  movel([0.215229, -1.349679, -2.570749, -0.791960, 1.570796, 1.786025],accel_mss,speed_ms,0,blend_radius_m)
  movel([0.214975, -1.350752, -2.570030, -0.791607, 1.570796, 1.785771],accel_mss,speed_ms,0,blend_radius_m)
  movel([0.216793, -1.350982, -2.569876, -0.791531, 1.570796, 1.787589],accel_mss,speed_ms,0,blend_radius_m)
  movel([0.217496, -1.351072, -2.569815, -0.791501, 1.570796, 1.788292],accel_mss,speed_ms,0,blend_radius_m)
  movel([0.218102, -1.351157, -2.569759, -0.791474, 1.570796, 1.788899],accel_mss,speed_ms,0,blend_radius_m)
  movel([0.218626, -1.351233, -2.569708, -0.791449, 1.570796, 1.789422],accel_mss,speed_ms,0,blend_radius_m)
  movel([0.218706, -1.351253, -2.569694, -0.791442, 1.570796, 1.789502],accel_mss,speed_ms,0,blend_radius_m)
  movel([0.218724, -1.351267, -2.569684, -0.791437, 1.570796, 1.789520],accel_mss,speed_ms,0,blend_radius_m)
  movel([0.218733, -1.351290, -2.569669, -0.791430, 1.570796, 1.789529],accel_mss,speed_ms,0,blend_radius_m)
  movel([0.218734, -1.351316, -2.569652, -0.791421, 1.570796, 1.789530],accel_mss,speed_ms,0,blend_radius_m)
  movel([0.218624, -1.351824, -2.569310, -0.791255, 1.570796, 1.789420],accel_mss,speed_ms,0,blend_radius_m)
  movel([0.218549, -1.352134, -2.569101, -0.791153, 1.570796, 1.789345],accel_mss,speed_ms,0,blend_radius_m)
  movel([0.218472, -1.352445, -2.568892, -0.791052, 1.570796, 1.789269],accel_mss,speed_ms,0,blend_radius_m)
  movel([0.218266, -1.353205, -2.568380, -0.790804, 1.570796, 1.789063],accel_mss,speed_ms,0,blend_radius_m)
  movel([0.216610, -1.359807, -2.563898, -0.788684, 1.570796, 1.787406],accel_mss,speed_ms,0,blend_radius_m)
  movel([0.214499, -1.360772, -2.563238, -0.788379, 1.570796, 1.785296],accel_mss,speed_ms,0,blend_radius_m)
  movel([0.212391, -1.361738, -2.562575, -0.788076, 1.570796, 1.783188],accel_mss,speed_ms,0,blend_radius_m)
  movel([0.212109, -1.362945, -2.561746, -0.787698, 1.570796, 1.782905],accel_mss,speed_ms,0,blend_radius_m)
  movel([0.211827, -1.364150, -2.560916, -0.787322, 1.570796, 1.782623],accel_mss,speed_ms,0,blend_radius_m)
  movel([0.210167, -1.364988, -2.560338, -0.787063, 1.570796, 1.780964],accel_mss,speed_ms,0,blend_radius_m)
  movel([0.208509, -1.365829, -2.559757, -0.786803, 1.570796, 1.779305],accel_mss,speed_ms,0,blend_radius_m)
  movel([0.208371, -1.366429, -2.559341, -0.786619, 1.570796, 1.779167],accel_mss,speed_ms,0,blend_radius_m)
  movel([0.208233, -1.367028, -2.558926, -0.786435, 1.570796, 1.779029],accel_mss,speed_ms,0,blend_radius_m)
  speed_ms = 0.003
  movel([0.208233, -1.370183, -2.560451, -0.781755, 1.570796, 1.779029],accel_mss,speed_ms,0,blend_radius_m)
  speed_ms = 0.007
  movel([0.192461, -1.373239, -2.558315, -0.780834, 1.570796, 1.763257],accel_mss,speed_ms,0,blend_radius_m)
  movel([0.176700, -1.376487, -2.556031, -0.779871, 1.570796, 1.747496],accel_mss,speed_ms,0,blend_radius_m)
  movel([0.177720, -1.375452, -2.556761, -0.780176, 1.570796, 1.748516],accel_mss,speed_ms,0,blend_radius_m)
  movel([0.178177, -1.374979, -2.557093, -0.780317, 1.570796, 1.748973],accel_mss,speed_ms,0,blend_radius_m)
  movel([0.178623, -1.374493, -2.557435, -0.780461, 1.570796, 1.749419],accel_mss,speed_ms,0,blend_radius_m)
  movel([0.179054, -1.374002, -2.557780, -0.780607, 1.570796, 1.749850],accel_mss,speed_ms,0,blend_radius_m)
  movel([0.179470, -1.373501, -2.558132, -0.780756, 1.570796, 1.750267],accel_mss,speed_ms,0,blend_radius_m)
  movel([0.179870, -1.372995, -2.558487, -0.780908, 1.570796, 1.750666],accel_mss,speed_ms,0,blend_radius_m)
  movel([0.180257, -1.372480, -2.558847, -0.781062, 1.570796, 1.751054],accel_mss,speed_ms,0,blend_radius_m)
  movel([0.180628, -1.371960, -2.559211, -0.781218, 1.570796, 1.751424],accel_mss,speed_ms,0,blend_radius_m)
  movel([0.180979, -1.371442, -2.559573, -0.781374, 1.570796, 1.751775],accel_mss,speed_ms,0,blend_radius_m)
  movel([0.181310, -1.370919, -2.559938, -0.781532, 1.570796, 1.752107],accel_mss,speed_ms,0,blend_radius_m)
  movel([0.181624, -1.370393, -2.560304, -0.781691, 1.570796, 1.752420],accel_mss,speed_ms,0,blend_radius_m)
  movel([0.181922, -1.369862, -2.560675, -0.781852, 1.570796, 1.752718],accel_mss,speed_ms,0,blend_radius_m)
  movel([0.182200, -1.369330, -2.561045, -0.782014, 1.570796, 1.752996],accel_mss,speed_ms,0,blend_radius_m)
  movel([0.182457, -1.368796, -2.561416, -0.782177, 1.570796, 1.753253],accel_mss,speed_ms,0,blend_radius_m)
  movel([0.182698, -1.368260, -2.561788, -0.782341, 1.570796, 1.753494],accel_mss,speed_ms,0,blend_radius_m)
  movel([0.182918, -1.367722, -2.562161, -0.782505, 1.570796, 1.753714],accel_mss,speed_ms,0,blend_radius_m)
  movel([0.183120, -1.367184, -2.562534, -0.782671, 1.570796, 1.753916],accel_mss,speed_ms,0,blend_radius_m)
  movel([0.183301, -1.366645, -2.562907, -0.782837, 1.570796, 1.754097],accel_mss,speed_ms,0,blend_radius_m)
  movel([0.183460, -1.366110, -2.563277, -0.783002, 1.570796, 1.754256],accel_mss,speed_ms,0,blend_radius_m)
  movel([0.183600, -1.365577, -2.563645, -0.783167, 1.570796, 1.754396],accel_mss,speed_ms,0,blend_radius_m)
  movel([0.183717, -1.365048, -2.564010, -0.783331, 1.570796, 1.754514],accel_mss,speed_ms,0,blend_radius_m)
  movel([0.183813, -1.364523, -2.564372, -0.783494, 1.570796, 1.754609],accel_mss,speed_ms,0,blend_radius_m)
  movel([0.183892, -1.363989, -2.564740, -0.783660, 1.570796, 1.754688],accel_mss,speed_ms,0,blend_radius_m)
  movel([0.183948, -1.363461, -2.565103, -0.783825, 1.570796, 1.754744],accel_mss,speed_ms,0,blend_radius_m)
  movel([0.183986, -1.362939, -2.565462, -0.783988, 1.570796, 1.754782],accel_mss,speed_ms,0,blend_radius_m)
  movel([0.184002, -1.362423, -2.565816, -0.784150, 1.570796, 1.754798],accel_mss,speed_ms,0,blend_radius_m)
  movel([0.183994, -1.361916, -2.566163, -0.784310, 1.570796, 1.754790],accel_mss,speed_ms,0,blend_radius_m)
  movel([0.183968, -1.361415, -2.566506, -0.784468, 1.570796, 1.754765],accel_mss,speed_ms,0,blend_radius_m)
  movel([0.183922, -1.360922, -2.566843, -0.784623, 1.570796, 1.754718],accel_mss,speed_ms,0,blend_radius_m)
  movel([0.183841, -1.360413, -2.567192, -0.784784, 1.570796, 1.754637],accel_mss,speed_ms,0,blend_radius_m)
  movel([0.183722, -1.359924, -2.567525, -0.784939, 1.570796, 1.754519],accel_mss,speed_ms,0,blend_radius_m)
  movel([0.183540, -1.359341, -2.567923, -0.785125, 1.570796, 1.754336],accel_mss,speed_ms,0,blend_radius_m)
  movel([0.183332, -1.358771, -2.568312, -0.785307, 1.570796, 1.754129],accel_mss,speed_ms,0,blend_radius_m)
  movel([0.183103, -1.358222, -2.568685, -0.785482, 1.570796, 1.753900],accel_mss,speed_ms,0,blend_radius_m)
  movel([0.182850, -1.357690, -2.569047, -0.785652, 1.570796, 1.753646],accel_mss,speed_ms,0,blend_radius_m)
  movel([0.182624, -1.357296, -2.569314, -0.785779, 1.570796, 1.753421],accel_mss,speed_ms,0,blend_radius_m)
  movel([0.182360, -1.356931, -2.569562, -0.785896, 1.570796, 1.753156],accel_mss,speed_ms,0,blend_radius_m)
  movel([0.181837, -1.356285, -2.570000, -0.786104, 1.570796, 1.752633],accel_mss,speed_ms,0,blend_radius_m)
  movel([0.183063, -1.355949, -2.570227, -0.786213, 1.570796, 1.753859],accel_mss,speed_ms,0,blend_radius_m)
  movel([0.183512, -1.355833, -2.570306, -0.786250, 1.570796, 1.754308],accel_mss,speed_ms,0,blend_radius_m)
  movel([0.183955, -1.355730, -2.570375, -0.786283, 1.570796, 1.754752],accel_mss,speed_ms,0,blend_radius_m)
  movel([0.188162, -1.354804, -2.571002, -0.786583, 1.570796, 1.758958],accel_mss,speed_ms,0,blend_radius_m)
  movel([0.193088, -1.353747, -2.571715, -0.786927, 1.570796, 1.763885],accel_mss,speed_ms,0,blend_radius_m)
  movel([0.198699, -1.352579, -2.572501, -0.787309, 1.570796, 1.769495],accel_mss,speed_ms,0,blend_radius_m)
  movel([0.213116, -1.349701, -2.574430, -0.788258, 1.570796, 1.783912],accel_mss,speed_ms,0,blend_radius_m)
  movel([0.212938, -1.350458, -2.573924, -0.788007, 1.570796, 1.783735],accel_mss,speed_ms,0,blend_radius_m)
  movel([0.212761, -1.351214, -2.573418, -0.787758, 1.570796, 1.783557],accel_mss,speed_ms,0,blend_radius_m)
  movel([0.213243, -1.351323, -2.573344, -0.787721, 1.570796, 1.784040],accel_mss,speed_ms,0,blend_radius_m)
  movel([0.215483, -1.351799, -2.573025, -0.787565, 1.570796, 1.786280],accel_mss,speed_ms,0,blend_radius_m)
  movel([0.215229, -1.352874, -2.572303, -0.787212, 1.570796, 1.786025],accel_mss,speed_ms,0,blend_radius_m)
  movel([0.214975, -1.353945, -2.571582, -0.786863, 1.570796, 1.785771],accel_mss,speed_ms,0,blend_radius_m)
  movel([0.216793, -1.354174, -2.571427, -0.786788, 1.570796, 1.787589],accel_mss,speed_ms,0,blend_radius_m)
  movel([0.217496, -1.354264, -2.571366, -0.786759, 1.570796, 1.788292],accel_mss,speed_ms,0,blend_radius_m)
  movel([0.218102, -1.354348, -2.571309, -0.786732, 1.570796, 1.788899],accel_mss,speed_ms,0,blend_radius_m)
  movel([0.218626, -1.354424, -2.571258, -0.786707, 1.570796, 1.789422],accel_mss,speed_ms,0,blend_radius_m)
  movel([0.218706, -1.354444, -2.571245, -0.786700, 1.570796, 1.789502],accel_mss,speed_ms,0,blend_radius_m)
  movel([0.218724, -1.354458, -2.571235, -0.786696, 1.570796, 1.789520],accel_mss,speed_ms,0,blend_radius_m)
  movel([0.218733, -1.354481, -2.571220, -0.786688, 1.570796, 1.789529],accel_mss,speed_ms,0,blend_radius_m)
  movel([0.218734, -1.354507, -2.571202, -0.786680, 1.570796, 1.789530],accel_mss,speed_ms,0,blend_radius_m)
  movel([0.218624, -1.355014, -2.570860, -0.786515, 1.570796, 1.789420],accel_mss,speed_ms,0,blend_radius_m)
  movel([0.218549, -1.355323, -2.570651, -0.786415, 1.570796, 1.789345],accel_mss,speed_ms,0,blend_radius_m)
  movel([0.218472, -1.355633, -2.570441, -0.786315, 1.570796, 1.789269],accel_mss,speed_ms,0,blend_radius_m)
  movel([0.218266, -1.356391, -2.569928, -0.786070, 1.570796, 1.789063],accel_mss,speed_ms,0,blend_radius_m)
  movel([0.216610, -1.362978, -2.565435, -0.783976, 1.570796, 1.787406],accel_mss,speed_ms,0,blend_radius_m)
  movel([0.214499, -1.363941, -2.564773, -0.783675, 1.570796, 1.785296],accel_mss,speed_ms,0,blend_radius_m)
  movel([0.212391, -1.364905, -2.564109, -0.783375, 1.570796, 1.783188],accel_mss,speed_ms,0,blend_radius_m)
  movel([0.212109, -1.366109, -2.563278, -0.783002, 1.570796, 1.782905],accel_mss,speed_ms,0,blend_radius_m)
  movel([0.211827, -1.367312, -2.562446, -0.782631, 1.570796, 1.782623],accel_mss,speed_ms,0,blend_radius_m)
  movel([0.210167, -1.368148, -2.561866, -0.782375, 1.570796, 1.780964],accel_mss,speed_ms,0,blend_radius_m)
  movel([0.208509, -1.368986, -2.561284, -0.782119, 1.570796, 1.779305],accel_mss,speed_ms,0,blend_radius_m)
  movel([0.208371, -1.369585, -2.560868, -0.781937, 1.570796, 1.779167],accel_mss,speed_ms,0,blend_radius_m)
  movel([0.208233, -1.370183, -2.560451, -0.781755, 1.570796, 1.779029],accel_mss,speed_ms,0,blend_radius_m)
  speed_ms = 0.003
  movel([0.208233, -1.357697, -2.554302, -0.800390, 1.570796, 1.779029],accel_mss,speed_ms,0,blend_radius_m)
  speed_ms = 0.01
  movel([0.208233, -1.333772, -2.541623, -0.836993, 1.570796, 1.779029],accel_mss,speed_ms,0,blend_radius_m)
  movel([0.180390, -1.333590, -2.541744, -0.837055, 1.570796, 1.751186],accel_mss,speed_ms,0,blend_radius_m)
  movel([0.180390, -1.357518, -2.554425, -0.800447, 1.570796, 1.751186],accel_mss,speed_ms,0,blend_radius_m)
  speed_ms = 0.003
  movel([0.180390, -1.366850, -2.559050, -0.786489, 1.570796, 1.751186],accel_mss,speed_ms,0,blend_radius_m)
  speed_ms = 0.007
  movel([0.180139, -1.367279, -2.558752, -0.786358, 1.570796, 1.750935],accel_mss,speed_ms,0,blend_radius_m)
  movel([0.179877, -1.367706, -2.558456, -0.786227, 1.570796, 1.750673],accel_mss,speed_ms,0,blend_radius_m)
  movel([0.179604, -1.368128, -2.558163, -0.786098, 1.570796, 1.750400],accel_mss,speed_ms,0,blend_radius_m)
  movel([0.179318, -1.368547, -2.557871, -0.785971, 1.570796, 1.750115],accel_mss,speed_ms,0,blend_radius_m)
  movel([0.179021, -1.368963, -2.557582, -0.785844, 1.570796, 1.749818],accel_mss,speed_ms,0,blend_radius_m)
  movel([0.178714, -1.369376, -2.557294, -0.785719, 1.570796, 1.749510],accel_mss,speed_ms,0,blend_radius_m)
  movel([0.178399, -1.369774, -2.557017, -0.785598, 1.570796, 1.749196],accel_mss,speed_ms,0,blend_radius_m)
  movel([0.178077, -1.370168, -2.556742, -0.785479, 1.570796, 1.748873],accel_mss,speed_ms,0,blend_radius_m)
  movel([0.177744, -1.370558, -2.556470, -0.785361, 1.570796, 1.748540],accel_mss,speed_ms,0,blend_radius_m)
  movel([0.177401, -1.370941, -2.556202, -0.785246, 1.570796, 1.748197],accel_mss,speed_ms,0,blend_radius_m)
  movel([0.177050, -1.371317, -2.555939, -0.785133, 1.570796, 1.747846],accel_mss,speed_ms,0,blend_radius_m)
  movel([0.176686, -1.371687, -2.555680, -0.785022, 1.570796, 1.747483],accel_mss,speed_ms,0,blend_radius_m)
  movel([0.176338, -1.372028, -2.555441, -0.784919, 1.570796, 1.747134],accel_mss,speed_ms,0,blend_radius_m)
  movel([0.175979, -1.372363, -2.555207, -0.784819, 1.570796, 1.746776],accel_mss,speed_ms,0,blend_radius_m)
  movel([0.175611, -1.372687, -2.554979, -0.784722, 1.570796, 1.746408],accel_mss,speed_ms,0,blend_radius_m)
  movel([0.175233, -1.373005, -2.554756, -0.784627, 1.570796, 1.746029],accel_mss,speed_ms,0,blend_radius_m)
  movel([0.174850, -1.373312, -2.554541, -0.784536, 1.570796, 1.745646],accel_mss,speed_ms,0,blend_radius_m)
  movel([0.174458, -1.373609, -2.554332, -0.784447, 1.570796, 1.745254],accel_mss,speed_ms,0,blend_radius_m)
  movel([0.174093, -1.373873, -2.554147, -0.784369, 1.570796, 1.744889],accel_mss,speed_ms,0,blend_radius_m)
  movel([0.173720, -1.374131, -2.553966, -0.784293, 1.570796, 1.744516],accel_mss,speed_ms,0,blend_radius_m)
  movel([0.173344, -1.374381, -2.553790, -0.784219, 1.570796, 1.744141],accel_mss,speed_ms,0,blend_radius_m)
  movel([0.172966, -1.374620, -2.553621, -0.784148, 1.570796, 1.743762],accel_mss,speed_ms,0,blend_radius_m)
  movel([0.172582, -1.374853, -2.553458, -0.784079, 1.570796, 1.743378],accel_mss,speed_ms,0,blend_radius_m)
  movel([0.172196, -1.375075, -2.553301, -0.784013, 1.570796, 1.742992],accel_mss,speed_ms,0,blend_radius_m)
  movel([0.171804, -1.375290, -2.553149, -0.783950, 1.570796, 1.742600],accel_mss,speed_ms,0,blend_radius_m)
  movel([0.171412, -1.375495, -2.553005, -0.783889, 1.570796, 1.742208],accel_mss,speed_ms,0,blend_radius_m)
  movel([0.171030, -1.375683, -2.552872, -0.783834, 1.570796, 1.741826],accel_mss,speed_ms,0,blend_radius_m)
  movel([0.170645, -1.375863, -2.552745, -0.783781, 1.570796, 1.741442],accel_mss,speed_ms,0,blend_radius_m)
  movel([0.170260, -1.376033, -2.552625, -0.783731, 1.570796, 1.741057],accel_mss,speed_ms,0,blend_radius_m)
  movel([0.169873, -1.376193, -2.552512, -0.783684, 1.570796, 1.740669],accel_mss,speed_ms,0,blend_radius_m)
  movel([0.169507, -1.376333, -2.552413, -0.783643, 1.570796, 1.740304],accel_mss,speed_ms,0,blend_radius_m)
  movel([0.169142, -1.376463, -2.552321, -0.783604, 1.570796, 1.739938],accel_mss,speed_ms,0,blend_radius_m)
  movel([0.168779, -1.376578, -2.552240, -0.783571, 1.570796, 1.739576],accel_mss,speed_ms,0,blend_radius_m)
  movel([0.168414, -1.376683, -2.552166, -0.783540, 1.570796, 1.739210],accel_mss,speed_ms,0,blend_radius_m)
  movel([0.167297, -1.376988, -2.551950, -0.783451, 1.570796, 1.738093],accel_mss,speed_ms,0,blend_radius_m)
  movel([0.168071, -1.372455, -2.555142, -0.784792, 1.570796, 1.738868],accel_mss,speed_ms,0,blend_radius_m)
  movel([0.168467, -1.370193, -2.556724, -0.785471, 1.570796, 1.739263],accel_mss,speed_ms,0,blend_radius_m)
  movel([0.169039, -1.367024, -2.558929, -0.786436, 1.570796, 1.739836],accel_mss,speed_ms,0,blend_radius_m)
  movel([0.169678, -1.363562, -2.561322, -0.787506, 1.570796, 1.740474],accel_mss,speed_ms,0,blend_radius_m)
  movel([0.170290, -1.360312, -2.563553, -0.788525, 1.570796, 1.741086],accel_mss,speed_ms,0,blend_radius_m)
  movel([0.171749, -1.352643, -2.568759, -0.790987, 1.570796, 1.742545],accel_mss,speed_ms,0,blend_radius_m)
  movel([0.172957, -1.352437, -2.568897, -0.791054, 1.570796, 1.743754],accel_mss,speed_ms,0,blend_radius_m)
  movel([0.173404, -1.352369, -2.568943, -0.791077, 1.570796, 1.744200],accel_mss,speed_ms,0,blend_radius_m)
  movel([0.173845, -1.352318, -2.568978, -0.791093, 1.570796, 1.744641],accel_mss,speed_ms,0,blend_radius_m)
  movel([0.174283, -1.352282, -2.569002, -0.791105, 1.570796, 1.745079],accel_mss,speed_ms,0,blend_radius_m)
  movel([0.174710, -1.352267, -2.569012, -0.791110, 1.570796, 1.745506],accel_mss,speed_ms,0,blend_radius_m)
  movel([0.175134, -1.352265, -2.569013, -0.791111, 1.570796, 1.745930],accel_mss,speed_ms,0,blend_radius_m)
  movel([0.175547, -1.352284, -2.569001, -0.791104, 1.570796, 1.746343],accel_mss,speed_ms,0,blend_radius_m)
  movel([0.175952, -1.352320, -2.568977, -0.791093, 1.570796, 1.746748],accel_mss,speed_ms,0,blend_radius_m)
  movel([0.176349, -1.352370, -2.568942, -0.791076, 1.570796, 1.747145],accel_mss,speed_ms,0,blend_radius_m)
  movel([0.176744, -1.352439, -2.568896, -0.791054, 1.570796, 1.747541],accel_mss,speed_ms,0,blend_radius_m)
  movel([0.177127, -1.352526, -2.568838, -0.791025, 1.570796, 1.747923],accel_mss,speed_ms,0,blend_radius_m)
  movel([0.177502, -1.352627, -2.568769, -0.790992, 1.570796, 1.748298],accel_mss,speed_ms,0,blend_radius_m)
  movel([0.177863, -1.352745, -2.568690, -0.790954, 1.570796, 1.748660],accel_mss,speed_ms,0,blend_radius_m)
  movel([0.178215, -1.352879, -2.568600, -0.790910, 1.570796, 1.749011],accel_mss,speed_ms,0,blend_radius_m)
  movel([0.178553, -1.353028, -2.568500, -0.790862, 1.570796, 1.749350],accel_mss,speed_ms,0,blend_radius_m)
  movel([0.178879, -1.353193, -2.568388, -0.790808, 1.570796, 1.749675],accel_mss,speed_ms,0,blend_radius_m)
  movel([0.179192, -1.353372, -2.568267, -0.790750, 1.570796, 1.749989],accel_mss,speed_ms,0,blend_radius_m)
  movel([0.179499, -1.353572, -2.568132, -0.790685, 1.570796, 1.750295],accel_mss,speed_ms,0,blend_radius_m)
  movel([0.179790, -1.353786, -2.567988, -0.790615, 1.570796, 1.750587],accel_mss,speed_ms,0,blend_radius_m)
  movel([0.180067, -1.354015, -2.567834, -0.790541, 1.570796, 1.750863],accel_mss,speed_ms,0,blend_radius_m)
  movel([0.180332, -1.354254, -2.567672, -0.790463, 1.570796, 1.751128],accel_mss,speed_ms,0,blend_radius_m)
  movel([0.180581, -1.354510, -2.567498, -0.790380, 1.570796, 1.751377],accel_mss,speed_ms,0,blend_radius_m)
  movel([0.180813, -1.354779, -2.567317, -0.790293, 1.570796, 1.751610],accel_mss,speed_ms,0,blend_radius_m)
  movel([0.181029, -1.355060, -2.567127, -0.790202, 1.570796, 1.751825],accel_mss,speed_ms,0,blend_radius_m)
  movel([0.181232, -1.355352, -2.566929, -0.790108, 1.570796, 1.752028],accel_mss,speed_ms,0,blend_radius_m)
  movel([0.181419, -1.355665, -2.566717, -0.790007, 1.570796, 1.752215],accel_mss,speed_ms,0,blend_radius_m)
  movel([0.181592, -1.355987, -2.566499, -0.789903, 1.570796, 1.752389],accel_mss,speed_ms,0,blend_radius_m)
  movel([0.181749, -1.356319, -2.566273, -0.789797, 1.570796, 1.752545],accel_mss,speed_ms,0,blend_radius_m)
  movel([0.181892, -1.356661, -2.566041, -0.789687, 1.570796, 1.752688],accel_mss,speed_ms,0,blend_radius_m)
  movel([0.182015, -1.357015, -2.565800, -0.789573, 1.570796, 1.752811],accel_mss,speed_ms,0,blend_radius_m)
  movel([0.182125, -1.357377, -2.565555, -0.789458, 1.570796, 1.752921],accel_mss,speed_ms,0,blend_radius_m)
  movel([0.182217, -1.357746, -2.565303, -0.789339, 1.570796, 1.753013],accel_mss,speed_ms,0,blend_radius_m)
  movel([0.182289, -1.358126, -2.565044, -0.789218, 1.570796, 1.753086],accel_mss,speed_ms,0,blend_radius_m)
  movel([0.182339, -1.358455, -2.564821, -0.789113, 1.570796, 1.753135],accel_mss,speed_ms,0,blend_radius_m)
  movel([0.182373, -1.358791, -2.564591, -0.789007, 1.570796, 1.753169],accel_mss,speed_ms,0,blend_radius_m)
  movel([0.182394, -1.359132, -2.564359, -0.788898, 1.570796, 1.753190],accel_mss,speed_ms,0,blend_radius_m)
  movel([0.182397, -1.359481, -2.564120, -0.788788, 1.570796, 1.753193],accel_mss,speed_ms,0,blend_radius_m)
  movel([0.182382, -1.360023, -2.563750, -0.788616, 1.570796, 1.753178],accel_mss,speed_ms,0,blend_radius_m)
  movel([0.182346, -1.360572, -2.563375, -0.788443, 1.570796, 1.753143],accel_mss,speed_ms,0,blend_radius_m)
  movel([0.182293, -1.361126, -2.562995, -0.788268, 1.570796, 1.753090],accel_mss,speed_ms,0,blend_radius_m)
  movel([0.182218, -1.361684, -2.562612, -0.788093, 1.570796, 1.753014],accel_mss,speed_ms,0,blend_radius_m)
  movel([0.182125, -1.362248, -2.562225, -0.787916, 1.570796, 1.752921],accel_mss,speed_ms,0,blend_radius_m)
  movel([0.182013, -1.362813, -2.561837, -0.787739, 1.570796, 1.752809],accel_mss,speed_ms,0,blend_radius_m)
  movel([0.181927, -1.363179, -2.561585, -0.787625, 1.570796, 1.752723],accel_mss,speed_ms,0,blend_radius_m)
  movel([0.181826, -1.363548, -2.561331, -0.787510, 1.570796, 1.752623],accel_mss,speed_ms,0,blend_radius_m)
  movel([0.181711, -1.363920, -2.561075, -0.787394, 1.570796, 1.752507],accel_mss,speed_ms,0,blend_radius_m)
  movel([0.181582, -1.364291, -2.560819, -0.787279, 1.570796, 1.752378],accel_mss,speed_ms,0,blend_radius_m)
  movel([0.181417, -1.364720, -2.560523, -0.787146, 1.570796, 1.752213],accel_mss,speed_ms,0,blend_radius_m)
  movel([0.181239, -1.365147, -2.560228, -0.787014, 1.570796, 1.752035],accel_mss,speed_ms,0,blend_radius_m)
  movel([0.181047, -1.365573, -2.559934, -0.786882, 1.570796, 1.751843],accel_mss,speed_ms,0,blend_radius_m)
  movel([0.180841, -1.366000, -2.559639, -0.786751, 1.570796, 1.751637],accel_mss,speed_ms,0,blend_radius_m)
  movel([0.180621, -1.366427, -2.559343, -0.786619, 1.570796, 1.751417],accel_mss,speed_ms,0,blend_radius_m)
  movel([0.180390, -1.366850, -2.559050, -0.786489, 1.570796, 1.751186],accel_mss,speed_ms,0,blend_radius_m)
  speed_ms = 0.003
  movel([0.180390, -1.370005, -2.560575, -0.781809, 1.570796, 1.751186],accel_mss,speed_ms,0,blend_radius_m)
  speed_ms = 0.007
  movel([0.180139, -1.370433, -2.560277, -0.781679, 1.570796, 1.750935],accel_mss,speed_ms,0,blend_radius_m)
  movel([0.179877, -1.370858, -2.559980, -0.781550, 1.570796, 1.750673],accel_mss,speed_ms,0,blend_radius_m)
  movel([0.179604, -1.371280, -2.559686, -0.781423, 1.570796, 1.750400],accel_mss,speed_ms,0,blend_radius_m)
  movel([0.179318, -1.371698, -2.559394, -0.781297, 1.570796, 1.750115],accel_mss,speed_ms,0,blend_radius_m)
  movel([0.179021, -1.372113, -2.559104, -0.781172, 1.570796, 1.749818],accel_mss,speed_ms,0,blend_radius_m)
  movel([0.178714, -1.372524, -2.558816, -0.781049, 1.570796, 1.749510],accel_mss,speed_ms,0,blend_radius_m)
  movel([0.178399, -1.372922, -2.558537, -0.780929, 1.570796, 1.749196],accel_mss,speed_ms,0,blend_radius_m)
  movel([0.178077, -1.373315, -2.558262, -0.780812, 1.570796, 1.748873],accel_mss,speed_ms,0,blend_radius_m)
  movel([0.177744, -1.373703, -2.557990, -0.780696, 1.570796, 1.748540],accel_mss,speed_ms,0,blend_radius_m)
  movel([0.177401, -1.374086, -2.557721, -0.780582, 1.570796, 1.748197],accel_mss,speed_ms,0,blend_radius_m)
  movel([0.177050, -1.374461, -2.557458, -0.780470, 1.570796, 1.747846],accel_mss,speed_ms,0,blend_radius_m)
  movel([0.176686, -1.374830, -2.557198, -0.780361, 1.570796, 1.747483],accel_mss,speed_ms,0,blend_radius_m)
  movel([0.176338, -1.375171, -2.556959, -0.780260, 1.570796, 1.747134],accel_mss,speed_ms,0,blend_radius_m)
  movel([0.175979, -1.375505, -2.556723, -0.780161, 1.570796, 1.746776],accel_mss,speed_ms,0,blend_radius_m)
  movel([0.175611, -1.375828, -2.556496, -0.780065, 1.570796, 1.746408],accel_mss,speed_ms,0,blend_radius_m)
  movel([0.175233, -1.376145, -2.556272, -0.779972, 1.570796, 1.746029],accel_mss,speed_ms,0,blend_radius_m)
  movel([0.174850, -1.376451, -2.556057, -0.779882, 1.570796, 1.745646],accel_mss,speed_ms,0,blend_radius_m)
  movel([0.174458, -1.376748, -2.555847, -0.779794, 1.570796, 1.745254],accel_mss,speed_ms,0,blend_radius_m)
  movel([0.174093, -1.377011, -2.555661, -0.779717, 1.570796, 1.744889],accel_mss,speed_ms,0,blend_radius_m)
  movel([0.173720, -1.377268, -2.555479, -0.779641, 1.570796, 1.744516],accel_mss,speed_ms,0,blend_radius_m)
  movel([0.173344, -1.377517, -2.555303, -0.779568, 1.570796, 1.744141],accel_mss,speed_ms,0,blend_radius_m)
  movel([0.172966, -1.377756, -2.555134, -0.779498, 1.570796, 1.743762],accel_mss,speed_ms,0,blend_radius_m)
  movel([0.172582, -1.377988, -2.554970, -0.779431, 1.570796, 1.743378],accel_mss,speed_ms,0,blend_radius_m)
  movel([0.172196, -1.378210, -2.554813, -0.779366, 1.570796, 1.742992],accel_mss,speed_ms,0,blend_radius_m)
  movel([0.171804, -1.378425, -2.554661, -0.779303, 1.570796, 1.742600],accel_mss,speed_ms,0,blend_radius_m)
  movel([0.171412, -1.378629, -2.554516, -0.779243, 1.570796, 1.742208],accel_mss,speed_ms,0,blend_radius_m)
  movel([0.171030, -1.378817, -2.554383, -0.779189, 1.570796, 1.741826],accel_mss,speed_ms,0,blend_radius_m)
  movel([0.170645, -1.378997, -2.554256, -0.779137, 1.570796, 1.741442],accel_mss,speed_ms,0,blend_radius_m)
  movel([0.170260, -1.379166, -2.554136, -0.779087, 1.570796, 1.741057],accel_mss,speed_ms,0,blend_radius_m)
  movel([0.169873, -1.379325, -2.554023, -0.779041, 1.570796, 1.740669],accel_mss,speed_ms,0,blend_radius_m)
  movel([0.169507, -1.379466, -2.553923, -0.779000, 1.570796, 1.740304],accel_mss,speed_ms,0,blend_radius_m)
  movel([0.169142, -1.379595, -2.553831, -0.778963, 1.570796, 1.739938],accel_mss,speed_ms,0,blend_radius_m)
  movel([0.168779, -1.379710, -2.553750, -0.778929, 1.570796, 1.739576],accel_mss,speed_ms,0,blend_radius_m)
  movel([0.168414, -1.379814, -2.553676, -0.778899, 1.570796, 1.739210],accel_mss,speed_ms,0,blend_radius_m)
  movel([0.167297, -1.380119, -2.553459, -0.778811, 1.570796, 1.738093],accel_mss,speed_ms,0,blend_radius_m)
  movel([0.168071, -1.375597, -2.556659, -0.780134, 1.570796, 1.738868],accel_mss,speed_ms,0,blend_radius_m)
  movel([0.168467, -1.373340, -2.558245, -0.780804, 1.570796, 1.739263],accel_mss,speed_ms,0,blend_radius_m)
  movel([0.169039, -1.370179, -2.560454, -0.781756, 1.570796, 1.739836],accel_mss,speed_ms,0,blend_radius_m)
  movel([0.169678, -1.366724, -2.562853, -0.782812, 1.570796, 1.740474],accel_mss,speed_ms,0,blend_radius_m)
  movel([0.170290, -1.363482, -2.565089, -0.783819, 1.570796, 1.741086],accel_mss,speed_ms,0,blend_radius_m)
  movel([0.171749, -1.355831, -2.570307, -0.786251, 1.570796, 1.742545],accel_mss,speed_ms,0,blend_radius_m)
  movel([0.172957, -1.355626, -2.570446, -0.786317, 1.570796, 1.743754],accel_mss,speed_ms,0,blend_radius_m)
  movel([0.173404, -1.355558, -2.570492, -0.786339, 1.570796, 1.744200],accel_mss,speed_ms,0,blend_radius_m)
  movel([0.173845, -1.355506, -2.570527, -0.786356, 1.570796, 1.744641],accel_mss,speed_ms,0,blend_radius_m)
  movel([0.174283, -1.355471, -2.570551, -0.786367, 1.570796, 1.745079],accel_mss,speed_ms,0,blend_radius_m)
  movel([0.174710, -1.355456, -2.570561, -0.786372, 1.570796, 1.745506],accel_mss,speed_ms,0,blend_radius_m)
  movel([0.175134, -1.355454, -2.570562, -0.786373, 1.570796, 1.745930],accel_mss,speed_ms,0,blend_radius_m)
  movel([0.175547, -1.355473, -2.570550, -0.786367, 1.570796, 1.746343],accel_mss,speed_ms,0,blend_radius_m)
  movel([0.175952, -1.355508, -2.570526, -0.786355, 1.570796, 1.746748],accel_mss,speed_ms,0,blend_radius_m)
  movel([0.176349, -1.355559, -2.570491, -0.786339, 1.570796, 1.747145],accel_mss,speed_ms,0,blend_radius_m)
  movel([0.176744, -1.355627, -2.570445, -0.786317, 1.570796, 1.747541],accel_mss,speed_ms,0,blend_radius_m)
  movel([0.177127, -1.355714, -2.570387, -0.786289, 1.570796, 1.747923],accel_mss,speed_ms,0,blend_radius_m)
  movel([0.177502, -1.355815, -2.570318, -0.786256, 1.570796, 1.748298],accel_mss,speed_ms,0,blend_radius_m)
  movel([0.177863, -1.355933, -2.570238, -0.786218, 1.570796, 1.748660],accel_mss,speed_ms,0,blend_radius_m)
  movel([0.178215, -1.356066, -2.570148, -0.786175, 1.570796, 1.749011],accel_mss,speed_ms,0,blend_radius_m)
  movel([0.178553, -1.356215, -2.570047, -0.786127, 1.570796, 1.749350],accel_mss,speed_ms,0,blend_radius_m)
  movel([0.178879, -1.356380, -2.569936, -0.786074, 1.570796, 1.749675],accel_mss,speed_ms,0,blend_radius_m)
  movel([0.179192, -1.356558, -2.569815, -0.786016, 1.570796, 1.749989],accel_mss,speed_ms,0,blend_radius_m)
  movel([0.179499, -1.356758, -2.569679, -0.785952, 1.570796, 1.750295],accel_mss,speed_ms,0,blend_radius_m)
  movel([0.179790, -1.356971, -2.569534, -0.785883, 1.570796, 1.750587],accel_mss,speed_ms,0,blend_radius_m)
  movel([0.180067, -1.357199, -2.569380, -0.785810, 1.570796, 1.750863],accel_mss,speed_ms,0,blend_radius_m)
  movel([0.180332, -1.357439, -2.569217, -0.785733, 1.570796, 1.751128],accel_mss,speed_ms,0,blend_radius_m)
  movel([0.180581, -1.357694, -2.569044, -0.785651, 1.570796, 1.751377],accel_mss,speed_ms,0,blend_radius_m)
  movel([0.180813, -1.357962, -2.568862, -0.785565, 1.570796, 1.751610],accel_mss,speed_ms,0,blend_radius_m)
  movel([0.181029, -1.358242, -2.568671, -0.785476, 1.570796, 1.751825],accel_mss,speed_ms,0,blend_radius_m)
  movel([0.181232, -1.358533, -2.568473, -0.785382, 1.570796, 1.752028],accel_mss,speed_ms,0,blend_radius_m)
  movel([0.181419, -1.358846, -2.568261, -0.785283, 1.570796, 1.752215],accel_mss,speed_ms,0,blend_radius_m)
  movel([0.181592, -1.359167, -2.568042, -0.785180, 1.570796, 1.752389],accel_mss,speed_ms,0,blend_radius_m)
  movel([0.181749, -1.359499, -2.567816, -0.785075, 1.570796, 1.752545],accel_mss,speed_ms,0,blend_radius_m)
  movel([0.181892, -1.359840, -2.567583, -0.784966, 1.570796, 1.752688],accel_mss,speed_ms,0,blend_radius_m)
  movel([0.182015, -1.360193, -2.567342, -0.784854, 1.570796, 1.752811],accel_mss,speed_ms,0,blend_radius_m)
  movel([0.182125, -1.360554, -2.567095, -0.784740, 1.570796, 1.752921],accel_mss,speed_ms,0,blend_radius_m)
  movel([0.182217, -1.360923, -2.566843, -0.784623, 1.570796, 1.753013],accel_mss,speed_ms,0,blend_radius_m)
  movel([0.182289, -1.361302, -2.566584, -0.784503, 1.570796, 1.753086],accel_mss,speed_ms,0,blend_radius_m)
  movel([0.182339, -1.361629, -2.566360, -0.784400, 1.570796, 1.753135],accel_mss,speed_ms,0,blend_radius_m)
  movel([0.182373, -1.361965, -2.566130, -0.784294, 1.570796, 1.753169],accel_mss,speed_ms,0,blend_radius_m)
  movel([0.182394, -1.362305, -2.565897, -0.784187, 1.570796, 1.753190],accel_mss,speed_ms,0,blend_radius_m)
  movel([0.182397, -1.362653, -2.565658, -0.784078, 1.570796, 1.753193],accel_mss,speed_ms,0,blend_radius_m)
  movel([0.182382, -1.363194, -2.565286, -0.783908, 1.570796, 1.753178],accel_mss,speed_ms,0,blend_radius_m)
  movel([0.182346, -1.363741, -2.564910, -0.783737, 1.570796, 1.753143],accel_mss,speed_ms,0,blend_radius_m)
  movel([0.182293, -1.364294, -2.564530, -0.783565, 1.570796, 1.753090],accel_mss,speed_ms,0,blend_radius_m)
  movel([0.182218, -1.364851, -2.564146, -0.783392, 1.570796, 1.753014],accel_mss,speed_ms,0,blend_radius_m)
  movel([0.182125, -1.365413, -2.563758, -0.783217, 1.570796, 1.752921],accel_mss,speed_ms,0,blend_radius_m)
  movel([0.182013, -1.365977, -2.563369, -0.783043, 1.570796, 1.752809],accel_mss,speed_ms,0,blend_radius_m)
  movel([0.181927, -1.366343, -2.563116, -0.782930, 1.570796, 1.752723],accel_mss,speed_ms,0,blend_radius_m)
  movel([0.181826, -1.366711, -2.562862, -0.782816, 1.570796, 1.752623],accel_mss,speed_ms,0,blend_radius_m)
  movel([0.181711, -1.367082, -2.562605, -0.782702, 1.570796, 1.752507],accel_mss,speed_ms,0,blend_radius_m)
  movel([0.181582, -1.367451, -2.562349, -0.782589, 1.570796, 1.752378],accel_mss,speed_ms,0,blend_radius_m)
  movel([0.181417, -1.367880, -2.562052, -0.782457, 1.570796, 1.752213],accel_mss,speed_ms,0,blend_radius_m)
  movel([0.181239, -1.368306, -2.561756, -0.782327, 1.570796, 1.752035],accel_mss,speed_ms,0,blend_radius_m)
  movel([0.181047, -1.368731, -2.561461, -0.782197, 1.570796, 1.751843],accel_mss,speed_ms,0,blend_radius_m)
  movel([0.180841, -1.369157, -2.561165, -0.782067, 1.570796, 1.751637],accel_mss,speed_ms,0,blend_radius_m)
  movel([0.180621, -1.369583, -2.560869, -0.781937, 1.570796, 1.751417],accel_mss,speed_ms,0,blend_radius_m)
  movel([0.180390, -1.370005, -2.560575, -0.781809, 1.570796, 1.751186],accel_mss,speed_ms,0,blend_radius_m)
  speed_ms = 0.003
  movel([0.180390, -1.357518, -2.554425, -0.800447, 1.570796, 1.751186],accel_mss,speed_ms,0,blend_radius_m)
  speed_ms = 0.01
  movel([0.180390, -1.333590, -2.541744, -0.837055, 1.570796, 1.751186],accel_mss,speed_ms,0,blend_radius_m)
  movel([0.171218, -1.350489, -2.530391, -0.831509, 1.570796, 1.742015],accel_mss,speed_ms,0,blend_radius_m)
  movel([0.171218, -1.374152, -2.542861, -0.795376, 1.570796, 1.742015],accel_mss,speed_ms,0,blend_radius_m)
  speed_ms = 0.003
  movel([0.171218, -1.383370, -2.547407, -0.781612, 1.570796, 1.742015],accel_mss,speed_ms,0,blend_radius_m)
  speed_ms = 0.007
  movel([0.171590, -1.383483, -2.547326, -0.781580, 1.570796, 1.742387],accel_mss,speed_ms,0,blend_radius_m)
  movel([0.171950, -1.383611, -2.547235, -0.781544, 1.570796, 1.742746],accel_mss,speed_ms,0,blend_radius_m)
  movel([0.172300, -1.383753, -2.547132, -0.781503, 1.570796, 1.743096],accel_mss,speed_ms,0,blend_radius_m)
  movel([0.172634, -1.383912, -2.547019, -0.781459, 1.570796, 1.743431],accel_mss,speed_ms,0,blend_radius_m)
  movel([0.172957, -1.384085, -2.546894, -0.781409, 1.570796, 1.743753],accel_mss,speed_ms,0,blend_radius_m)
  movel([0.173267, -1.384274, -2.546759, -0.781356, 1.570796, 1.744064],accel_mss,speed_ms,0,blend_radius_m)
  movel([0.173560, -1.384479, -2.546612, -0.781298, 1.570796, 1.744357],accel_mss,speed_ms,0,blend_radius_m)
  movel([0.173841, -1.384697, -2.546455, -0.781237, 1.570796, 1.744638],accel_mss,speed_ms,0,blend_radius_m)
  movel([0.174108, -1.384930, -2.546288, -0.781171, 1.570796, 1.744904],accel_mss,speed_ms,0,blend_radius_m)
  movel([0.174357, -1.385178, -2.546110, -0.781102, 1.570796, 1.745154],accel_mss,speed_ms,0,blend_radius_m)
  movel([0.174598, -1.385446, -2.545917, -0.781026, 1.570796, 1.745394],accel_mss,speed_ms,0,blend_radius_m)
  movel([0.174827, -1.385726, -2.545715, -0.780948, 1.570796, 1.745623],accel_mss,speed_ms,0,blend_radius_m)
  movel([0.175037, -1.386019, -2.545504, -0.780866, 1.570796, 1.745834],accel_mss,speed_ms,0,blend_radius_m)
  movel([0.175231, -1.386326, -2.545283, -0.780780, 1.570796, 1.746027],accel_mss,speed_ms,0,blend_radius_m)
  movel([0.175408, -1.386642, -2.545055, -0.780691, 1.570796, 1.746205],accel_mss,speed_ms,0,blend_radius_m)
  movel([0.175569, -1.386972, -2.544817, -0.780599, 1.570796, 1.746365],accel_mss,speed_ms,0,blend_radius_m)
  movel([0.175712, -1.387310, -2.544573, -0.780505, 1.570796, 1.746509],accel_mss,speed_ms,0,blend_radius_m)
  movel([0.175837, -1.387660, -2.544321, -0.780408, 1.570796, 1.746633],accel_mss,speed_ms,0,blend_radius_m)
  movel([0.175945, -1.388019, -2.544061, -0.780309, 1.570796, 1.746742],accel_mss,speed_ms,0,blend_radius_m)
  movel([0.176036, -1.388388, -2.543795, -0.780207, 1.570796, 1.746832],accel_mss,speed_ms,0,blend_radius_m)
  movel([0.176114, -1.388774, -2.543515, -0.780100, 1.570796, 1.746910],accel_mss,speed_ms,0,blend_radius_m)
  movel([0.176171, -1.389170, -2.543228, -0.779991, 1.570796, 1.746967],accel_mss,speed_ms,0,blend_radius_m)
  movel([0.176214, -1.389571, -2.542938, -0.779881, 1.570796, 1.747010],accel_mss,speed_ms,0,blend_radius_m)
  movel([0.176241, -1.389979, -2.542642, -0.779769, 1.570796, 1.747037],accel_mss,speed_ms,0,blend_radius_m)
  movel([0.176248, -1.390395, -2.542339, -0.779655, 1.570796, 1.747044],accel_mss,speed_ms,0,blend_radius_m)
  movel([0.176241, -1.390816, -2.542034, -0.779539, 1.570796, 1.747037],accel_mss,speed_ms,0,blend_radius_m)
  movel([0.176216, -1.391242, -2.541724, -0.779423, 1.570796, 1.747012],accel_mss,speed_ms,0,blend_radius_m)
  movel([0.176175, -1.391672, -2.541411, -0.779306, 1.570796, 1.746971],accel_mss,speed_ms,0,blend_radius_m)
  movel([0.176116, -1.392109, -2.541093, -0.779188, 1.570796, 1.746912],accel_mss,speed_ms,0,blend_radius_m)
  movel([0.176041, -1.392547, -2.540773, -0.779069, 1.570796, 1.746837],accel_mss,speed_ms,0,blend_radius_m)
  movel([0.175989, -1.392809, -2.540582, -0.778998, 1.570796, 1.746785],accel_mss,speed_ms,0,blend_radius_m)
  movel([0.175927, -1.393072, -2.540390, -0.778927, 1.570796, 1.746724],accel_mss,speed_ms,0,blend_radius_m)
  movel([0.175855, -1.393369, -2.540173, -0.778847, 1.570796, 1.746651],accel_mss,speed_ms,0,blend_radius_m)
  movel([0.175776, -1.393667, -2.539955, -0.778767, 1.570796, 1.746572],accel_mss,speed_ms,0,blend_radius_m)
  movel([0.175696, -1.393953, -2.539746, -0.778690, 1.570796, 1.746493],accel_mss,speed_ms,0,blend_radius_m)
  movel([0.175610, -1.394240, -2.539536, -0.778613, 1.570796, 1.746406],accel_mss,speed_ms,0,blend_radius_m)
  movel([0.175538, -1.394464, -2.539372, -0.778553, 1.570796, 1.746335],accel_mss,speed_ms,0,blend_radius_m)
  movel([0.175458, -1.394688, -2.539208, -0.778493, 1.570796, 1.746254],accel_mss,speed_ms,0,blend_radius_m)
  movel([0.175287, -1.395126, -2.538887, -0.778376, 1.570796, 1.746083],accel_mss,speed_ms,0,blend_radius_m)
  movel([0.175101, -1.395562, -2.538567, -0.778260, 1.570796, 1.745897],accel_mss,speed_ms,0,blend_radius_m)
  movel([0.174901, -1.395999, -2.538247, -0.778144, 1.570796, 1.745697],accel_mss,speed_ms,0,blend_radius_m)
  movel([0.174688, -1.396434, -2.537927, -0.778028, 1.570796, 1.745484],accel_mss,speed_ms,0,blend_radius_m)
  movel([0.174461, -1.396867, -2.537609, -0.777913, 1.570796, 1.745258],accel_mss,speed_ms,0,blend_radius_m)
  movel([0.174219, -1.397299, -2.537291, -0.777799, 1.570796, 1.745016],accel_mss,speed_ms,0,blend_radius_m)
  movel([0.173967, -1.397727, -2.536975, -0.777686, 1.570796, 1.744763],accel_mss,speed_ms,0,blend_radius_m)
  movel([0.173701, -1.398156, -2.536660, -0.777574, 1.570796, 1.744497],accel_mss,speed_ms,0,blend_radius_m)
  movel([0.173423, -1.398578, -2.536348, -0.777463, 1.570796, 1.744219],accel_mss,speed_ms,0,blend_radius_m)
  movel([0.173144, -1.398980, -2.536051, -0.777358, 1.570796, 1.743940],accel_mss,speed_ms,0,blend_radius_m)
  movel([0.172850, -1.399379, -2.535756, -0.777254, 1.570796, 1.743647],accel_mss,speed_ms,0,blend_radius_m)
  movel([0.172544, -1.399772, -2.535466, -0.777151, 1.570796, 1.743341],accel_mss,speed_ms,0,blend_radius_m)
  movel([0.172228, -1.400161, -2.535178, -0.777050, 1.570796, 1.743024],accel_mss,speed_ms,0,blend_radius_m)
  movel([0.171900, -1.400542, -2.534896, -0.776951, 1.570796, 1.742696],accel_mss,speed_ms,0,blend_radius_m)
  movel([0.171559, -1.400919, -2.534616, -0.776854, 1.570796, 1.742355],accel_mss,speed_ms,0,blend_radius_m)
  movel([0.171209, -1.401288, -2.534343, -0.776759, 1.570796, 1.742005],accel_mss,speed_ms,0,blend_radius_m)
  movel([0.170849, -1.401648, -2.534075, -0.776666, 1.570796, 1.741645],accel_mss,speed_ms,0,blend_radius_m)
  movel([0.170477, -1.402001, -2.533813, -0.776575, 1.570796, 1.741273],accel_mss,speed_ms,0,blend_radius_m)
  movel([0.170106, -1.402339, -2.533562, -0.776488, 1.570796, 1.740902],accel_mss,speed_ms,0,blend_radius_m)
  movel([0.169725, -1.402667, -2.533318, -0.776404, 1.570796, 1.740522],accel_mss,speed_ms,0,blend_radius_m)
  movel([0.169338, -1.402986, -2.533080, -0.776322, 1.570796, 1.740134],accel_mss,speed_ms,0,blend_radius_m)
  movel([0.168941, -1.403295, -2.532850, -0.776243, 1.570796, 1.739738],accel_mss,speed_ms,0,blend_radius_m)
  movel([0.168540, -1.403593, -2.532629, -0.776168, 1.570796, 1.739337],accel_mss,speed_ms,0,blend_radius_m)
  movel([0.168130, -1.403882, -2.532413, -0.776094, 1.570796, 1.738926],accel_mss,speed_ms,0,blend_radius_m)
  movel([0.167713, -1.404161, -2.532205, -0.776023, 1.570796, 1.738509],accel_mss,speed_ms,0,blend_radius_m)
  movel([0.167293, -1.404428, -2.532006, -0.775955, 1.570796, 1.738089],accel_mss,speed_ms,0,blend_radius_m)
  movel([0.166867, -1.404682, -2.531816, -0.775891, 1.570796, 1.737663],accel_mss,speed_ms,0,blend_radius_m)
  movel([0.166434, -1.404925, -2.531634, -0.775829, 1.570796, 1.737231],accel_mss,speed_ms,0,blend_radius_m)
  movel([0.165997, -1.405157, -2.531461, -0.775771, 1.570796, 1.736793],accel_mss,speed_ms,0,blend_radius_m)
  movel([0.165557, -1.405378, -2.531296, -0.775715, 1.570796, 1.736354],accel_mss,speed_ms,0,blend_radius_m)
  movel([0.165116, -1.405585, -2.531141, -0.775663, 1.570796, 1.735912],accel_mss,speed_ms,0,blend_radius_m)
  movel([0.164673, -1.405778, -2.530996, -0.775614, 1.570796, 1.735469],accel_mss,speed_ms,0,blend_radius_m)
  movel([0.164228, -1.405958, -2.530862, -0.775569, 1.570796, 1.735024],accel_mss,speed_ms,0,blend_radius_m)
  movel([0.163781, -1.406126, -2.530736, -0.775527, 1.570796, 1.734577],accel_mss,speed_ms,0,blend_radius_m)
  movel([0.163334, -1.406280, -2.530621, -0.775488, 1.570796, 1.734130],accel_mss,speed_ms,0,blend_radius_m)
  movel([0.162890, -1.406419, -2.530516, -0.775453, 1.570796, 1.733686],accel_mss,speed_ms,0,blend_radius_m)
  movel([0.162475, -1.406539, -2.530427, -0.775423, 1.570796, 1.733271],accel_mss,speed_ms,0,blend_radius_m)
  movel([0.162111, -1.406633, -2.530356, -0.775400, 1.570796, 1.732908],accel_mss,speed_ms,0,blend_radius_m)
  movel([0.161806, -1.406708, -2.530300, -0.775381, 1.570796, 1.732602],accel_mss,speed_ms,0,blend_radius_m)
  movel([0.161769, -1.406711, -2.530297, -0.775380, 1.570796, 1.732565],accel_mss,speed_ms,0,blend_radius_m)
  movel([0.161734, -1.406704, -2.530303, -0.775382, 1.570796, 1.732531],accel_mss,speed_ms,0,blend_radius_m)
  movel([0.161716, -1.406692, -2.530312, -0.775385, 1.570796, 1.732512],accel_mss,speed_ms,0,blend_radius_m)
  movel([0.161706, -1.406672, -2.530327, -0.775390, 1.570796, 1.732503],accel_mss,speed_ms,0,blend_radius_m)
  movel([0.161706, -1.406648, -2.530345, -0.775396, 1.570796, 1.732502],accel_mss,speed_ms,0,blend_radius_m)
  movel([0.162290, -1.403310, -2.532840, -0.776240, 1.570796, 1.733086],accel_mss,speed_ms,0,blend_radius_m)
  movel([0.162618, -1.401449, -2.534223, -0.776717, 1.570796, 1.733414],accel_mss,speed_ms,0,blend_radius_m)
  movel([0.162952, -1.399581, -2.535607, -0.777201, 1.570796, 1.733748],accel_mss,speed_ms,0,blend_radius_m)
  movel([0.163765, -1.395132, -2.538883, -0.778374, 1.570796, 1.734561],accel_mss,speed_ms,0,blend_radius_m)
  movel([0.165943, -1.383394, -2.547390, -0.781605, 1.570796, 1.736739],accel_mss,speed_ms,0,blend_radius_m)
  movel([0.167049, -1.383219, -2.547516, -0.781655, 1.570796, 1.737845],accel_mss,speed_ms,0,blend_radius_m)
  movel([0.167499, -1.383155, -2.547561, -0.781673, 1.570796, 1.738295],accel_mss,speed_ms,0,blend_radius_m)
  movel([0.167941, -1.383111, -2.547592, -0.781685, 1.570796, 1.738737],accel_mss,speed_ms,0,blend_radius_m)
  movel([0.168380, -1.383081, -2.547614, -0.781694, 1.570796, 1.739176],accel_mss,speed_ms,0,blend_radius_m)
  movel([0.168810, -1.383072, -2.547620, -0.781697, 1.570796, 1.739607],accel_mss,speed_ms,0,blend_radius_m)
  movel([0.169236, -1.383079, -2.547616, -0.781695, 1.570796, 1.740032],accel_mss,speed_ms,0,blend_radius_m)
  movel([0.169650, -1.383102, -2.547599, -0.781688, 1.570796, 1.740447],accel_mss,speed_ms,0,blend_radius_m)
  movel([0.170057, -1.383144, -2.547569, -0.781676, 1.570796, 1.740853],accel_mss,speed_ms,0,blend_radius_m)
  movel([0.170454, -1.383201, -2.547528, -0.781660, 1.570796, 1.741250],accel_mss,speed_ms,0,blend_radius_m)
  movel([0.170843, -1.383277, -2.547474, -0.781638, 1.570796, 1.741639],accel_mss,speed_ms,0,blend_radius_m)
  movel([0.171218, -1.383370, -2.547407, -0.781612, 1.570796, 1.742015],accel_mss,speed_ms,0,blend_radius_m)
  speed_ms = 0.003
  movel([0.171218, -1.386485, -2.548906, -0.776998, 1.570796, 1.742015],accel_mss,speed_ms,0,blend_radius_m)
  speed_ms = 0.007
  movel([0.171590, -1.386597, -2.548825, -0.776966, 1.570796, 1.742387],accel_mss,speed_ms,0,blend_radius_m)
  movel([0.171950, -1.386725, -2.548733, -0.776931, 1.570796, 1.742746],accel_mss,speed_ms,0,blend_radius_m)
  movel([0.172300, -1.386867, -2.548631, -0.776891, 1.570796, 1.743096],accel_mss,speed_ms,0,blend_radius_m)
  movel([0.172634, -1.387025, -2.548517, -0.776847, 1.570796, 1.743431],accel_mss,speed_ms,0,blend_radius_m)
  movel([0.172957, -1.387198, -2.548392, -0.776798, 1.570796, 1.743753],accel_mss,speed_ms,0,blend_radius_m)
  movel([0.173267, -1.387387, -2.548256, -0.776746, 1.570796, 1.744064],accel_mss,speed_ms,0,blend_radius_m)
  movel([0.173560, -1.387591, -2.548109, -0.776689, 1.570796, 1.744357],accel_mss,speed_ms,0,blend_radius_m)
  movel([0.173841, -1.387808, -2.547952, -0.776628, 1.570796, 1.744638],accel_mss,speed_ms,0,blend_radius_m)
  movel([0.174108, -1.388041, -2.547784, -0.776563, 1.570796, 1.744904],accel_mss,speed_ms,0,blend_radius_m)
  movel([0.174357, -1.388288, -2.547606, -0.776495, 1.570796, 1.745154],accel_mss,speed_ms,0,blend_radius_m)
  movel([0.174598, -1.388555, -2.547413, -0.776421, 1.570796, 1.745394],accel_mss,speed_ms,0,blend_radius_m)
  movel([0.174827, -1.388836, -2.547210, -0.776343, 1.570796, 1.745623],accel_mss,speed_ms,0,blend_radius_m)
  movel([0.175037, -1.389128, -2.546999, -0.776262, 1.570796, 1.745834],accel_mss,speed_ms,0,blend_radius_m)
  movel([0.175231, -1.389434, -2.546777, -0.776178, 1.570796, 1.746027],accel_mss,speed_ms,0,blend_radius_m)
  movel([0.175408, -1.389749, -2.546549, -0.776091, 1.570796, 1.746205],accel_mss,speed_ms,0,blend_radius_m)
  movel([0.175569, -1.390078, -2.546311, -0.776000, 1.570796, 1.746365],accel_mss,speed_ms,0,blend_radius_m)
  movel([0.175712, -1.390415, -2.546066, -0.775907, 1.570796, 1.746509],accel_mss,speed_ms,0,blend_radius_m)
  movel([0.175837, -1.390764, -2.545813, -0.775812, 1.570796, 1.746633],accel_mss,speed_ms,0,blend_radius_m)
  movel([0.175945, -1.391122, -2.545553, -0.775714, 1.570796, 1.746742],accel_mss,speed_ms,0,blend_radius_m)
  movel([0.176036, -1.391490, -2.545286, -0.775613, 1.570796, 1.746832],accel_mss,speed_ms,0,blend_radius_m)
  movel([0.176114, -1.391875, -2.545006, -0.775508, 1.570796, 1.746910],accel_mss,speed_ms,0,blend_radius_m)
  movel([0.176171, -1.392270, -2.544718, -0.775400, 1.570796, 1.746967],accel_mss,speed_ms,0,blend_radius_m)
  movel([0.176214, -1.392671, -2.544427, -0.775292, 1.570796, 1.747010],accel_mss,speed_ms,0,blend_radius_m)
  movel([0.176241, -1.393078, -2.544130, -0.775181, 1.570796, 1.747037],accel_mss,speed_ms,0,blend_radius_m)
  movel([0.176248, -1.393493, -2.543827, -0.775069, 1.570796, 1.747044],accel_mss,speed_ms,0,blend_radius_m)
  movel([0.176241, -1.393913, -2.543521, -0.774956, 1.570796, 1.747037],accel_mss,speed_ms,0,blend_radius_m)
  movel([0.176216, -1.394338, -2.543210, -0.774841, 1.570796, 1.747012],accel_mss,speed_ms,0,blend_radius_m)
  movel([0.176175, -1.394766, -2.542897, -0.774726, 1.570796, 1.746971],accel_mss,speed_ms,0,blend_radius_m)
  movel([0.176116, -1.395202, -2.542578, -0.774609, 1.570796, 1.746912],accel_mss,speed_ms,0,blend_radius_m)
  movel([0.176041, -1.395639, -2.542258, -0.774492, 1.570796, 1.746837],accel_mss,speed_ms,0,blend_radius_m)
  movel([0.175989, -1.395900, -2.542066, -0.774422, 1.570796, 1.746785],accel_mss,speed_ms,0,blend_radius_m)
  movel([0.175927, -1.396163, -2.541873, -0.774352, 1.570796, 1.746724],accel_mss,speed_ms,0,blend_radius_m)
  movel([0.175855, -1.396459, -2.541656, -0.774273, 1.570796, 1.746651],accel_mss,speed_ms,0,blend_radius_m)
  movel([0.175776, -1.396757, -2.541438, -0.774194, 1.570796, 1.746572],accel_mss,speed_ms,0,blend_radius_m)
  movel([0.175696, -1.397042, -2.541228, -0.774119, 1.570796, 1.746493],accel_mss,speed_ms,0,blend_radius_m)
  movel([0.175610, -1.397328, -2.541018, -0.774043, 1.570796, 1.746406],accel_mss,speed_ms,0,blend_radius_m)
  movel([0.175538, -1.397552, -2.540853, -0.773984, 1.570796, 1.746335],accel_mss,speed_ms,0,blend_radius_m)
  movel([0.175458, -1.397775, -2.540689, -0.773925, 1.570796, 1.746254],accel_mss,speed_ms,0,blend_radius_m)
  movel([0.175287, -1.398212, -2.540368, -0.773810, 1.570796, 1.746083],accel_mss,speed_ms,0,blend_radius_m)
  movel([0.175101, -1.398647, -2.540047, -0.773695, 1.570796, 1.745897],accel_mss,speed_ms,0,blend_radius_m)
  movel([0.174901, -1.399082, -2.539726, -0.773581, 1.570796, 1.745697],accel_mss,speed_ms,0,blend_radius_m)
  movel([0.174688, -1.399516, -2.539406, -0.773467, 1.570796, 1.745484],accel_mss,speed_ms,0,blend_radius_m)
  movel([0.174461, -1.399949, -2.539086, -0.773354, 1.570796, 1.745258],accel_mss,speed_ms,0,blend_radius_m)
  movel([0.174219, -1.400380, -2.538768, -0.773242, 1.570796, 1.745016],accel_mss,speed_ms,0,blend_radius_m)
  movel([0.173967, -1.400807, -2.538452, -0.773131, 1.570796, 1.744763],accel_mss,speed_ms,0,blend_radius_m)
  movel([0.173701, -1.401234, -2.538135, -0.773020, 1.570796, 1.744497],accel_mss,speed_ms,0,blend_radius_m)
  movel([0.173423, -1.401655, -2.537823, -0.772911, 1.570796, 1.744219],accel_mss,speed_ms,0,blend_radius_m)
  movel([0.173144, -1.402056, -2.537525, -0.772807, 1.570796, 1.743940],accel_mss,speed_ms,0,blend_radius_m)
  movel([0.172850, -1.402454, -2.537230, -0.772705, 1.570796, 1.743647],accel_mss,speed_ms,0,blend_radius_m)
  movel([0.172544, -1.402846, -2.536939, -0.772604, 1.570796, 1.743341],accel_mss,speed_ms,0,blend_radius_m)
  movel([0.172228, -1.403234, -2.536650, -0.772505, 1.570796, 1.743024],accel_mss,speed_ms,0,blend_radius_m)
  movel([0.171900, -1.403614, -2.536368, -0.772407, 1.570796, 1.742696],accel_mss,speed_ms,0,blend_radius_m)
  movel([0.171559, -1.403990, -2.536087, -0.772311, 1.570796, 1.742355],accel_mss,speed_ms,0,blend_radius_m)
  movel([0.171209, -1.404358, -2.535813, -0.772217, 1.570796, 1.742005],accel_mss,speed_ms,0,blend_radius_m)
  movel([0.170849, -1.404718, -2.535545, -0.772126, 1.570796, 1.741645],accel_mss,speed_ms,0,blend_radius_m)
  movel([0.170477, -1.405070, -2.535283, -0.772037, 1.570796, 1.741273],accel_mss,speed_ms,0,blend_radius_m)
  movel([0.170106, -1.405407, -2.535031, -0.771951, 1.570796, 1.740902],accel_mss,speed_ms,0,blend_radius_m)
  movel([0.169725, -1.405734, -2.534786, -0.771868, 1.570796, 1.740522],accel_mss,speed_ms,0,blend_radius_m)
  movel([0.169338, -1.406053, -2.534548, -0.771788, 1.570796, 1.740134],accel_mss,speed_ms,0,blend_radius_m)
  movel([0.168941, -1.406361, -2.534318, -0.771711, 1.570796, 1.739738],accel_mss,speed_ms,0,blend_radius_m)
  movel([0.168540, -1.406657, -2.534096, -0.771636, 1.570796, 1.739337],accel_mss,speed_ms,0,blend_radius_m)
  movel([0.168130, -1.406946, -2.533879, -0.771563, 1.570796, 1.738926],accel_mss,speed_ms,0,blend_radius_m)
  movel([0.167713, -1.407224, -2.533671, -0.771494, 1.570796, 1.738509],accel_mss,speed_ms,0,blend_radius_m)
  movel([0.167293, -1.407490, -2.533472, -0.771427, 1.570796, 1.738089],accel_mss,speed_ms,0,blend_radius_m)
  movel([0.166867, -1.407744, -2.533281, -0.771364, 1.570796, 1.737663],accel_mss,speed_ms,0,blend_radius_m)
  movel([0.166434, -1.407986, -2.533099, -0.771303, 1.570796, 1.737231],accel_mss,speed_ms,0,blend_radius_m)
  movel([0.165997, -1.408218, -2.532925, -0.771246, 1.570796, 1.736793],accel_mss,speed_ms,0,blend_radius_m)
  movel([0.165557, -1.408438, -2.532760, -0.771191, 1.570796, 1.736354],accel_mss,speed_ms,0,blend_radius_m)
  movel([0.165116, -1.408645, -2.532605, -0.771139, 1.570796, 1.735912],accel_mss,speed_ms,0,blend_radius_m)
  movel([0.164673, -1.408837, -2.532460, -0.771092, 1.570796, 1.735469],accel_mss,speed_ms,0,blend_radius_m)
  movel([0.164228, -1.409017, -2.532325, -0.771047, 1.570796, 1.735024],accel_mss,speed_ms,0,blend_radius_m)
  movel([0.163781, -1.409184, -2.532199, -0.771006, 1.570796, 1.734577],accel_mss,speed_ms,0,blend_radius_m)
  movel([0.163334, -1.409338, -2.532083, -0.770968, 1.570796, 1.734130],accel_mss,speed_ms,0,blend_radius_m)
  movel([0.162890, -1.409477, -2.531979, -0.770933, 1.570796, 1.733686],accel_mss,speed_ms,0,blend_radius_m)
  movel([0.162475, -1.409596, -2.531889, -0.770904, 1.570796, 1.733271],accel_mss,speed_ms,0,blend_radius_m)
  movel([0.162111, -1.409690, -2.531818, -0.770881, 1.570796, 1.732908],accel_mss,speed_ms,0,blend_radius_m)
  movel([0.161806, -1.409764, -2.531762, -0.770862, 1.570796, 1.732602],accel_mss,speed_ms,0,blend_radius_m)
  movel([0.161769, -1.409768, -2.531760, -0.770861, 1.570796, 1.732565],accel_mss,speed_ms,0,blend_radius_m)
  movel([0.161734, -1.409761, -2.531765, -0.770863, 1.570796, 1.732531],accel_mss,speed_ms,0,blend_radius_m)
  movel([0.161716, -1.409749, -2.531774, -0.770866, 1.570796, 1.732512],accel_mss,speed_ms,0,blend_radius_m)
  movel([0.161706, -1.409729, -2.531789, -0.770871, 1.570796, 1.732503],accel_mss,speed_ms,0,blend_radius_m)
  movel([0.161706, -1.409705, -2.531807, -0.770877, 1.570796, 1.732502],accel_mss,speed_ms,0,blend_radius_m)
  movel([0.162290, -1.406375, -2.534307, -0.771707, 1.570796, 1.733086],accel_mss,speed_ms,0,blend_radius_m)
  movel([0.162618, -1.404519, -2.535694, -0.772177, 1.570796, 1.733414],accel_mss,speed_ms,0,blend_radius_m)
  movel([0.162952, -1.402656, -2.537080, -0.772653, 1.570796, 1.733748],accel_mss,speed_ms,0,blend_radius_m)
  movel([0.163765, -1.398218, -2.540363, -0.773808, 1.570796, 1.734561],accel_mss,speed_ms,0,blend_radius_m)
  movel([0.165943, -1.386509, -2.548889, -0.776991, 1.570796, 1.736739],accel_mss,speed_ms,0,blend_radius_m)
  movel([0.167049, -1.386334, -2.549015, -0.777040, 1.570796, 1.737845],accel_mss,speed_ms,0,blend_radius_m)
  movel([0.167499, -1.386270, -2.549061, -0.777058, 1.570796, 1.738295],accel_mss,speed_ms,0,blend_radius_m)
  movel([0.167941, -1.386227, -2.549092, -0.777070, 1.570796, 1.738737],accel_mss,speed_ms,0,blend_radius_m)
  movel([0.168380, -1.386197, -2.549113, -0.777079, 1.570796, 1.739176],accel_mss,speed_ms,0,blend_radius_m)
  movel([0.168810, -1.386188, -2.549120, -0.777081, 1.570796, 1.739607],accel_mss,speed_ms,0,blend_radius_m)
  movel([0.169236, -1.386194, -2.549115, -0.777079, 1.570796, 1.740032],accel_mss,speed_ms,0,blend_radius_m)
  movel([0.169650, -1.386218, -2.549098, -0.777073, 1.570796, 1.740447],accel_mss,speed_ms,0,blend_radius_m)
  movel([0.170057, -1.386260, -2.549068, -0.777061, 1.570796, 1.740853],accel_mss,speed_ms,0,blend_radius_m)
  movel([0.170454, -1.386317, -2.549027, -0.777045, 1.570796, 1.741250],accel_mss,speed_ms,0,blend_radius_m)
  movel([0.170843, -1.386392, -2.548973, -0.777024, 1.570796, 1.741639],accel_mss,speed_ms,0,blend_radius_m)
  movel([0.171218, -1.386485, -2.548906, -0.776998, 1.570796, 1.742015],accel_mss,speed_ms,0,blend_radius_m)
  speed_ms = 0.003
  movel([0.171218, -1.374152, -2.542861, -0.795376, 1.570796, 1.742015],accel_mss,speed_ms,0,blend_radius_m)
  speed_ms = 0.01
  movel([0.171218, -1.350489, -2.530391, -0.831509, 1.570796, 1.742015],accel_mss,speed_ms,0,blend_radius_m)
  movel([0.293421, -1.317023, -2.552513, -0.842853, 1.570796, 1.864217],accel_mss,speed_ms,0,blend_radius_m)
  movel([0.293421, -1.341199, -2.565402, -0.805788, 1.570796, 1.864217],accel_mss,speed_ms,0,blend_radius_m)
  speed_ms = 0.003
  movel([0.293421, -1.350639, -2.570106, -0.791644, 1.570796, 1.864217],accel_mss,speed_ms,0,blend_radius_m)
  speed_ms = 0.007
  movel([0.293458, -1.350455, -2.570229, -0.791704, 1.570796, 1.864254],accel_mss,speed_ms,0,blend_radius_m)
  movel([0.293505, -1.350268, -2.570355, -0.791766, 1.570796, 1.864301],accel_mss,speed_ms,0,blend_radius_m)
  movel([0.293560, -1.350079, -2.570481, -0.791828, 1.570796, 1.864356],accel_mss,speed_ms,0,blend_radius_m)
  movel([0.293625, -1.349890, -2.570608, -0.791891, 1.570796, 1.864421],accel_mss,speed_ms,0,blend_radius_m)
  movel([0.293697, -1.349699, -2.570736, -0.791954, 1.570796, 1.864493],accel_mss,speed_ms,0,blend_radius_m)
  movel([0.293778, -1.349510, -2.570863, -0.792016, 1.570796, 1.864574],accel_mss,speed_ms,0,blend_radius_m)
  movel([0.293942, -1.349162, -2.571096, -0.792131, 1.570796, 1.864738],accel_mss,speed_ms,0,blend_radius_m)
  movel([0.294118, -1.348813, -2.571329, -0.792247, 1.570796, 1.864914],accel_mss,speed_ms,0,blend_radius_m)
  movel([0.294299, -1.348485, -2.571548, -0.792356, 1.570796, 1.865096],accel_mss,speed_ms,0,blend_radius_m)
  movel([0.294494, -1.348160, -2.571765, -0.792464, 1.570796, 1.865290],accel_mss,speed_ms,0,blend_radius_m)
  movel([0.294707, -1.347837, -2.571980, -0.792571, 1.570796, 1.865503],accel_mss,speed_ms,0,blend_radius_m)
  movel([0.294935, -1.347519, -2.572192, -0.792677, 1.570796, 1.865731],accel_mss,speed_ms,0,blend_radius_m)
  movel([0.295171, -1.347214, -2.572396, -0.792779, 1.570796, 1.865967],accel_mss,speed_ms,0,blend_radius_m)
  movel([0.295421, -1.346913, -2.572596, -0.792879, 1.570796, 1.866218],accel_mss,speed_ms,0,blend_radius_m)
  movel([0.295683, -1.346623, -2.572790, -0.792977, 1.570796, 1.866480],accel_mss,speed_ms,0,blend_radius_m)
  movel([0.295960, -1.346339, -2.572978, -0.793072, 1.570796, 1.866756],accel_mss,speed_ms,0,blend_radius_m)
  movel([0.296244, -1.346068, -2.573158, -0.793162, 1.570796, 1.867040],accel_mss,speed_ms,0,blend_radius_m)
  movel([0.296539, -1.345807, -2.573332, -0.793250, 1.570796, 1.867336],accel_mss,speed_ms,0,blend_radius_m)
  movel([0.296842, -1.345559, -2.573497, -0.793333, 1.570796, 1.867639],accel_mss,speed_ms,0,blend_radius_m)
  movel([0.297156, -1.345323, -2.573654, -0.793413, 1.570796, 1.867952],accel_mss,speed_ms,0,blend_radius_m)
  movel([0.297478, -1.345097, -2.573803, -0.793489, 1.570796, 1.868274],accel_mss,speed_ms,0,blend_radius_m)
  movel([0.297805, -1.344886, -2.573943, -0.793560, 1.570796, 1.868601],accel_mss,speed_ms,0,blend_radius_m)
  movel([0.298137, -1.344689, -2.574074, -0.793626, 1.570796, 1.868934],accel_mss,speed_ms,0,blend_radius_m)
  movel([0.298476, -1.344508, -2.574194, -0.793687, 1.570796, 1.869272],accel_mss,speed_ms,0,blend_radius_m)
  movel([0.298814, -1.344337, -2.574307, -0.793745, 1.570796, 1.869610],accel_mss,speed_ms,0,blend_radius_m)
  movel([0.299154, -1.344175, -2.574414, -0.793800, 1.570796, 1.869950],accel_mss,speed_ms,0,blend_radius_m)
  movel([0.299297, -1.344111, -2.574457, -0.793821, 1.570796, 1.870094],accel_mss,speed_ms,0,blend_radius_m)
  movel([0.299437, -1.344058, -2.574492, -0.793839, 1.570796, 1.870233],accel_mss,speed_ms,0,blend_radius_m)
  movel([0.299579, -1.344012, -2.574522, -0.793855, 1.570796, 1.870376],accel_mss,speed_ms,0,blend_radius_m)
  movel([0.299806, -1.343954, -2.574561, -0.793874, 1.570796, 1.870602],accel_mss,speed_ms,0,blend_radius_m)
  movel([0.300029, -1.343912, -2.574589, -0.793889, 1.570796, 1.870826],accel_mss,speed_ms,0,blend_radius_m)
  movel([0.300440, -1.343855, -2.574626, -0.793908, 1.570796, 1.871236],accel_mss,speed_ms,0,blend_radius_m)
  movel([0.300848, -1.343806, -2.574659, -0.793924, 1.570796, 1.871644],accel_mss,speed_ms,0,blend_radius_m)
  movel([0.301256, -1.343761, -2.574689, -0.793940, 1.570796, 1.872053],accel_mss,speed_ms,0,blend_radius_m)
  movel([0.301660, -1.343723, -2.574713, -0.793952, 1.570796, 1.872457],accel_mss,speed_ms,0,blend_radius_m)
  movel([0.301873, -1.343715, -2.574719, -0.793955, 1.570796, 1.872670],accel_mss,speed_ms,0,blend_radius_m)
  movel([0.302078, -1.343723, -2.574713, -0.793952, 1.570796, 1.872875],accel_mss,speed_ms,0,blend_radius_m)
  movel([0.302201, -1.343739, -2.574703, -0.793947, 1.570796, 1.872997],accel_mss,speed_ms,0,blend_radius_m)
  movel([0.302316, -1.343762, -2.574688, -0.793939, 1.570796, 1.873112],accel_mss,speed_ms,0,blend_radius_m)
  movel([0.302428, -1.343797, -2.574665, -0.793928, 1.570796, 1.873224],accel_mss,speed_ms,0,blend_radius_m)
  movel([0.302685, -1.343890, -2.574603, -0.793896, 1.570796, 1.873482],accel_mss,speed_ms,0,blend_radius_m)
  movel([0.302935, -1.343993, -2.574535, -0.793861, 1.570796, 1.873731],accel_mss,speed_ms,0,blend_radius_m)
  movel([0.303162, -1.344099, -2.574465, -0.793825, 1.570796, 1.873959],accel_mss,speed_ms,0,blend_radius_m)
  movel([0.303378, -1.344220, -2.574385, -0.793784, 1.570796, 1.874174],accel_mss,speed_ms,0,blend_radius_m)
  movel([0.303581, -1.344356, -2.574295, -0.793739, 1.570796, 1.874378],accel_mss,speed_ms,0,blend_radius_m)
  movel([0.303769, -1.344505, -2.574196, -0.793688, 1.570796, 1.874565],accel_mss,speed_ms,0,blend_radius_m)
  movel([0.303943, -1.344665, -2.574090, -0.793634, 1.570796, 1.874739],accel_mss,speed_ms,0,blend_radius_m)
  movel([0.304101, -1.344840, -2.573974, -0.793575, 1.570796, 1.874897],accel_mss,speed_ms,0,blend_radius_m)
  movel([0.304243, -1.345026, -2.573851, -0.793513, 1.570796, 1.875039],accel_mss,speed_ms,0,blend_radius_m)
  movel([0.304372, -1.345222, -2.573720, -0.793446, 1.570796, 1.875168],accel_mss,speed_ms,0,blend_radius_m)
  movel([0.304484, -1.345434, -2.573580, -0.793375, 1.570796, 1.875280],accel_mss,speed_ms,0,blend_radius_m)
  movel([0.304578, -1.345657, -2.573431, -0.793300, 1.570796, 1.875375],accel_mss,speed_ms,0,blend_radius_m)
  movel([0.304660, -1.345891, -2.573276, -0.793222, 1.570796, 1.875456],accel_mss,speed_ms,0,blend_radius_m)
  movel([0.304722, -1.346133, -2.573115, -0.793141, 1.570796, 1.875518],accel_mss,speed_ms,0,blend_radius_m)
  movel([0.304772, -1.346390, -2.572944, -0.793055, 1.570796, 1.875569],accel_mss,speed_ms,0,blend_radius_m)
  movel([0.304805, -1.346656, -2.572768, -0.792966, 1.570796, 1.875602],accel_mss,speed_ms,0,blend_radius_m)
  movel([0.304821, -1.346930, -2.572585, -0.792874, 1.570796, 1.875618],accel_mss,speed_ms,0,blend_radius_m)
  movel([0.304822, -1.347208, -2.572400, -0.792781, 1.570796, 1.875619],accel_mss,speed_ms,0,blend_radius_m)
  movel([0.304810, -1.347440, -2.572245, -0.792704, 1.570796, 1.875606],accel_mss,speed_ms,0,blend_radius_m)
  movel([0.304780, -1.347676, -2.572088, -0.792625, 1.570796, 1.875576],accel_mss,speed_ms,0,blend_radius_m)
  movel([0.304736, -1.347919, -2.571926, -0.792544, 1.570796, 1.875532],accel_mss,speed_ms,0,blend_radius_m)
  movel([0.304671, -1.348208, -2.571733, -0.792448, 1.570796, 1.875468],accel_mss,speed_ms,0,blend_radius_m)
  movel([0.304594, -1.348501, -2.571537, -0.792351, 1.570796, 1.875391],accel_mss,speed_ms,0,blend_radius_m)
  movel([0.304507, -1.348797, -2.571339, -0.792252, 1.570796, 1.875303],accel_mss,speed_ms,0,blend_radius_m)
  movel([0.304411, -1.349090, -2.571144, -0.792155, 1.570796, 1.875208],accel_mss,speed_ms,0,blend_radius_m)
  movel([0.304305, -1.349386, -2.570946, -0.792057, 1.570796, 1.875102],accel_mss,speed_ms,0,blend_radius_m)
  movel([0.304190, -1.349680, -2.570749, -0.791960, 1.570796, 1.874987],accel_mss,speed_ms,0,blend_radius_m)
  movel([0.304083, -1.349922, -2.570587, -0.791880, 1.570796, 1.874879],accel_mss,speed_ms,0,blend_radius_m)
  movel([0.303962, -1.350165, -2.570424, -0.791800, 1.570796, 1.874758],accel_mss,speed_ms,0,blend_radius_m)
  movel([0.303829, -1.350404, -2.570264, -0.791721, 1.570796, 1.874626],accel_mss,speed_ms,0,blend_radius_m)
  movel([0.303632, -1.350727, -2.570047, -0.791615, 1.570796, 1.874429],accel_mss,speed_ms,0,blend_radius_m)
  movel([0.303419, -1.351046, -2.569833, -0.791510, 1.570796, 1.874215],accel_mss,speed_ms,0,blend_radius_m)
  movel([0.303192, -1.351358, -2.569623, -0.791408, 1.570796, 1.873989],accel_mss,speed_ms,0,blend_radius_m)
  movel([0.302951, -1.351668, -2.569415, -0.791306, 1.570796, 1.873747],accel_mss,speed_ms,0,blend_radius_m)
  movel([0.302696, -1.351970, -2.569212, -0.791207, 1.570796, 1.873492],accel_mss,speed_ms,0,blend_radius_m)
  movel([0.302434, -1.352257, -2.569019, -0.791113, 1.570796, 1.873230],accel_mss,speed_ms,0,blend_radius_m)
  movel([0.302161, -1.352536, -2.568831, -0.791022, 1.570796, 1.872957],accel_mss,speed_ms,0,blend_radius_m)
  movel([0.301874, -1.352806, -2.568649, -0.790934, 1.570796, 1.872671],accel_mss,speed_ms,0,blend_radius_m)
  movel([0.301579, -1.353067, -2.568473, -0.790849, 1.570796, 1.872375],accel_mss,speed_ms,0,blend_radius_m)
  movel([0.301274, -1.353316, -2.568305, -0.790768, 1.570796, 1.872070],accel_mss,speed_ms,0,blend_radius_m)
  movel([0.300964, -1.353549, -2.568148, -0.790692, 1.570796, 1.871761],accel_mss,speed_ms,0,blend_radius_m)
  movel([0.300645, -1.353771, -2.567998, -0.790620, 1.570796, 1.871441],accel_mss,speed_ms,0,blend_radius_m)
  movel([0.300323, -1.353979, -2.567858, -0.790552, 1.570796, 1.871119],accel_mss,speed_ms,0,blend_radius_m)
  movel([0.299992, -1.354172, -2.567727, -0.790490, 1.570796, 1.870788],accel_mss,speed_ms,0,blend_radius_m)
  movel([0.299659, -1.354351, -2.567607, -0.790432, 1.570796, 1.870455],accel_mss,speed_ms,0,blend_radius_m)
  movel([0.299323, -1.354516, -2.567495, -0.790378, 1.570796, 1.870119],accel_mss,speed_ms,0,blend_radius_m)
  movel([0.298983, -1.354665, -2.567394, -0.790330, 1.570796, 1.869779],accel_mss,speed_ms,0,blend_radius_m)
  movel([0.298641, -1.354798, -2.567304, -0.790287, 1.570796, 1.869437],accel_mss,speed_ms,0,blend_radius_m)
  movel([0.298303, -1.354912, -2.567227, -0.790250, 1.570796, 1.869100],accel_mss,speed_ms,0,blend_radius_m)
  movel([0.297963, -1.355013, -2.567159, -0.790218, 1.570796, 1.868759],accel_mss,speed_ms,0,blend_radius_m)
  movel([0.297675, -1.355081, -2.567112, -0.790196, 1.570796, 1.868471],accel_mss,speed_ms,0,blend_radius_m)
  movel([0.297387, -1.355134, -2.567077, -0.790179, 1.570796, 1.868183],accel_mss,speed_ms,0,blend_radius_m)
  movel([0.297107, -1.355170, -2.567052, -0.790167, 1.570796, 1.867903],accel_mss,speed_ms,0,blend_radius_m)
  movel([0.296830, -1.355190, -2.567038, -0.790160, 1.570796, 1.867626],accel_mss,speed_ms,0,blend_radius_m)
  movel([0.296563, -1.355192, -2.567037, -0.790160, 1.570796, 1.867359],accel_mss,speed_ms,0,blend_radius_m)
  movel([0.296302, -1.355177, -2.567047, -0.790164, 1.570796, 1.867098],accel_mss,speed_ms,0,blend_radius_m)
  movel([0.296048, -1.355146, -2.567068, -0.790175, 1.570796, 1.866844],accel_mss,speed_ms,0,blend_radius_m)
  movel([0.295793, -1.355095, -2.567103, -0.790191, 1.570796, 1.866589],accel_mss,speed_ms,0,blend_radius_m)
  movel([0.295549, -1.355031, -2.567146, -0.790212, 1.570796, 1.866346],accel_mss,speed_ms,0,blend_radius_m)
  movel([0.295313, -1.354952, -2.567200, -0.790237, 1.570796, 1.866110],accel_mss,speed_ms,0,blend_radius_m)
  movel([0.295089, -1.354857, -2.567264, -0.790268, 1.570796, 1.865885],accel_mss,speed_ms,0,blend_radius_m)
  movel([0.294878, -1.354748, -2.567338, -0.790303, 1.570796, 1.865675],accel_mss,speed_ms,0,blend_radius_m)
  movel([0.294679, -1.354626, -2.567421, -0.790343, 1.570796, 1.865475],accel_mss,speed_ms,0,blend_radius_m)
  movel([0.294491, -1.354489, -2.567513, -0.790387, 1.570796, 1.865287],accel_mss,speed_ms,0,blend_radius_m)
  movel([0.294312, -1.354331, -2.567620, -0.790438, 1.570796, 1.865108],accel_mss,speed_ms,0,blend_radius_m)
  movel([0.294143, -1.354164, -2.567733, -0.790492, 1.570796, 1.864940],accel_mss,speed_ms,0,blend_radius_m)
  movel([0.293991, -1.353980, -2.567857, -0.790552, 1.570796, 1.864787],accel_mss,speed_ms,0,blend_radius_m)
  movel([0.293854, -1.353787, -2.567988, -0.790615, 1.570796, 1.864650],accel_mss,speed_ms,0,blend_radius_m)
  movel([0.293731, -1.353582, -2.568126, -0.790681, 1.570796, 1.864528],accel_mss,speed_ms,0,blend_radius_m)
  movel([0.293624, -1.353367, -2.568271, -0.790751, 1.570796, 1.864420],accel_mss,speed_ms,0,blend_radius_m)
  movel([0.293532, -1.353141, -2.568423, -0.790825, 1.570796, 1.864328],accel_mss,speed_ms,0,blend_radius_m)
  movel([0.293455, -1.352901, -2.568585, -0.790903, 1.570796, 1.864252],accel_mss,speed_ms,0,blend_radius_m)
  movel([0.293393, -1.352654, -2.568752, -0.790984, 1.570796, 1.864189],accel_mss,speed_ms,0,blend_radius_m)
  movel([0.293350, -1.352397, -2.568924, -0.791067, 1.570796, 1.864146],accel_mss,speed_ms,0,blend_radius_m)
  movel([0.293321, -1.352134, -2.569101, -0.791153, 1.570796, 1.864117],accel_mss,speed_ms,0,blend_radius_m)
  movel([0.293308, -1.351863, -2.569284, -0.791242, 1.570796, 1.864105],accel_mss,speed_ms,0,blend_radius_m)
  movel([0.293312, -1.351584, -2.569471, -0.791333, 1.570796, 1.864108],accel_mss,speed_ms,0,blend_radius_m)
  movel([0.293331, -1.351302, -2.569661, -0.791426, 1.570796, 1.864127],accel_mss,speed_ms,0,blend_radius_m)
  movel([0.293369, -1.350972, -2.569882, -0.791534, 1.570796, 1.864165],accel_mss,speed_ms,0,blend_radius_m)
  movel([0.293421, -1.350639, -2.570106, -0.791644, 1.570796, 1.864217],accel_mss,speed_ms,0,blend_radius_m)
  speed_ms = 0.003
  movel([0.293421, -1.353831, -2.571658, -0.786900, 1.570796, 1.864217],accel_mss,speed_ms,0,blend_radius_m)
  speed_ms = 0.007
  movel([0.293458, -1.353648, -2.571781, -0.786960, 1.570796, 1.864254],accel_mss,speed_ms,0,blend_radius_m)
  movel([0.293505, -1.353461, -2.571907, -0.787021, 1.570796, 1.864301],accel_mss,speed_ms,0,blend_radius_m)
  movel([0.293560, -1.353273, -2.572034, -0.787082, 1.570796, 1.864356],accel_mss,speed_ms,0,blend_radius_m)
  movel([0.293625, -1.353084, -2.572161, -0.787144, 1.570796, 1.864421],accel_mss,speed_ms,0,blend_radius_m)
  movel([0.293697, -1.352894, -2.572289, -0.787206, 1.570796, 1.864493],accel_mss,speed_ms,0,blend_radius_m)
  movel([0.293778, -1.352705, -2.572416, -0.787268, 1.570796, 1.864574],accel_mss,speed_ms,0,blend_radius_m)
  movel([0.293942, -1.352358, -2.572650, -0.787381, 1.570796, 1.864738],accel_mss,speed_ms,0,blend_radius_m)
  movel([0.294118, -1.352009, -2.572884, -0.787496, 1.570796, 1.864914],accel_mss,speed_ms,0,blend_radius_m)
  movel([0.294299, -1.351682, -2.573103, -0.787603, 1.570796, 1.865096],accel_mss,speed_ms,0,blend_radius_m)
  movel([0.294494, -1.351358, -2.573321, -0.787710, 1.570796, 1.865290],accel_mss,speed_ms,0,blend_radius_m)
  movel([0.294707, -1.351036, -2.573537, -0.787816, 1.570796, 1.865503],accel_mss,speed_ms,0,blend_radius_m)
  movel([0.294935, -1.350719, -2.573749, -0.787921, 1.570796, 1.865731],accel_mss,speed_ms,0,blend_radius_m)
  movel([0.295171, -1.350414, -2.573953, -0.788021, 1.570796, 1.865967],accel_mss,speed_ms,0,blend_radius_m)
  movel([0.295421, -1.350114, -2.574154, -0.788121, 1.570796, 1.866218],accel_mss,speed_ms,0,blend_radius_m)
  movel([0.295683, -1.349824, -2.574348, -0.788217, 1.570796, 1.866480],accel_mss,speed_ms,0,blend_radius_m)
  movel([0.295960, -1.349542, -2.574537, -0.788311, 1.570796, 1.866756],accel_mss,speed_ms,0,blend_radius_m)
  movel([0.296244, -1.349271, -2.574717, -0.788400, 1.570796, 1.867040],accel_mss,speed_ms,0,blend_radius_m)
  movel([0.296539, -1.349011, -2.574891, -0.788487, 1.570796, 1.867336],accel_mss,speed_ms,0,blend_radius_m)
  movel([0.296842, -1.348763, -2.575057, -0.788569, 1.570796, 1.867639],accel_mss,speed_ms,0,blend_radius_m)
  movel([0.297156, -1.348527, -2.575214, -0.788648, 1.570796, 1.867952],accel_mss,speed_ms,0,blend_radius_m)
  movel([0.297478, -1.348302, -2.575364, -0.788723, 1.570796, 1.868274],accel_mss,speed_ms,0,blend_radius_m)
  movel([0.297805, -1.348092, -2.575504, -0.788793, 1.570796, 1.868601],accel_mss,speed_ms,0,blend_radius_m)
  movel([0.298137, -1.347895, -2.575635, -0.788859, 1.570796, 1.868934],accel_mss,speed_ms,0,blend_radius_m)
  movel([0.298476, -1.347715, -2.575755, -0.788919, 1.570796, 1.869272],accel_mss,speed_ms,0,blend_radius_m)
  movel([0.298814, -1.347544, -2.575869, -0.788976, 1.570796, 1.869610],accel_mss,speed_ms,0,blend_radius_m)
  movel([0.299154, -1.347382, -2.575977, -0.789030, 1.570796, 1.869950],accel_mss,speed_ms,0,blend_radius_m)
  movel([0.299297, -1.347318, -2.576019, -0.789052, 1.570796, 1.870094],accel_mss,speed_ms,0,blend_radius_m)
  movel([0.299437, -1.347266, -2.576054, -0.789069, 1.570796, 1.870233],accel_mss,speed_ms,0,blend_radius_m)
  movel([0.299579, -1.347220, -2.576085, -0.789085, 1.570796, 1.870376],accel_mss,speed_ms,0,blend_radius_m)
  movel([0.299806, -1.347161, -2.576123, -0.789104, 1.570796, 1.870602],accel_mss,speed_ms,0,blend_radius_m)
  movel([0.300029, -1.347120, -2.576151, -0.789118, 1.570796, 1.870826],accel_mss,speed_ms,0,blend_radius_m)
  movel([0.300440, -1.347063, -2.576189, -0.789137, 1.570796, 1.871236],accel_mss,speed_ms,0,blend_radius_m)
  movel([0.300848, -1.347014, -2.576222, -0.789154, 1.570796, 1.871644],accel_mss,speed_ms,0,blend_radius_m)
  movel([0.301256, -1.346969, -2.576251, -0.789169, 1.570796, 1.872053],accel_mss,speed_ms,0,blend_radius_m)
  movel([0.301660, -1.346932, -2.576276, -0.789181, 1.570796, 1.872457],accel_mss,speed_ms,0,blend_radius_m)
  movel([0.301873, -1.346923, -2.576282, -0.789184, 1.570796, 1.872670],accel_mss,speed_ms,0,blend_radius_m)
  movel([0.302078, -1.346931, -2.576276, -0.789181, 1.570796, 1.872875],accel_mss,speed_ms,0,blend_radius_m)
  movel([0.302201, -1.346947, -2.576266, -0.789176, 1.570796, 1.872997],accel_mss,speed_ms,0,blend_radius_m)
  movel([0.302316, -1.346970, -2.576251, -0.789168, 1.570796, 1.873112],accel_mss,speed_ms,0,blend_radius_m)
  movel([0.302428, -1.347005, -2.576228, -0.789157, 1.570796, 1.873224],accel_mss,speed_ms,0,blend_radius_m)
  movel([0.302685, -1.347098, -2.576166, -0.789125, 1.570796, 1.873482],accel_mss,speed_ms,0,blend_radius_m)
  movel([0.302935, -1.347201, -2.576097, -0.789091, 1.570796, 1.873731],accel_mss,speed_ms,0,blend_radius_m)
  movel([0.303162, -1.347306, -2.576027, -0.789056, 1.570796, 1.873959],accel_mss,speed_ms,0,blend_radius_m)
  movel([0.303378, -1.347427, -2.575947, -0.789015, 1.570796, 1.874174],accel_mss,speed_ms,0,blend_radius_m)
  movel([0.303581, -1.347563, -2.575856, -0.788970, 1.570796, 1.874378],accel_mss,speed_ms,0,blend_radius_m)
  movel([0.303769, -1.347711, -2.575757, -0.788920, 1.570796, 1.874565],accel_mss,speed_ms,0,blend_radius_m)
  movel([0.303943, -1.347871, -2.575651, -0.788867, 1.570796, 1.874739],accel_mss,speed_ms,0,blend_radius_m)
  movel([0.304101, -1.348046, -2.575535, -0.788808, 1.570796, 1.874897],accel_mss,speed_ms,0,blend_radius_m)
  movel([0.304243, -1.348231, -2.575411, -0.788747, 1.570796, 1.875039],accel_mss,speed_ms,0,blend_radius_m)
  movel([0.304372, -1.348427, -2.575281, -0.788681, 1.570796, 1.875168],accel_mss,speed_ms,0,blend_radius_m)
  movel([0.304484, -1.348639, -2.575140, -0.788611, 1.570796, 1.875280],accel_mss,speed_ms,0,blend_radius_m)
  movel([0.304578, -1.348861, -2.574991, -0.788537, 1.570796, 1.875375],accel_mss,speed_ms,0,blend_radius_m)
  movel([0.304660, -1.349094, -2.574836, -0.788459, 1.570796, 1.875456],accel_mss,speed_ms,0,blend_radius_m)
  movel([0.304722, -1.349336, -2.574674, -0.788379, 1.570796, 1.875518],accel_mss,speed_ms,0,blend_radius_m)
  movel([0.304772, -1.349592, -2.574503, -0.788294, 1.570796, 1.875569],accel_mss,speed_ms,0,blend_radius_m)
  movel([0.304805, -1.349857, -2.574326, -0.788206, 1.570796, 1.875602],accel_mss,speed_ms,0,blend_radius_m)
  movel([0.304821, -1.350131, -2.574143, -0.788115, 1.570796, 1.875618],accel_mss,speed_ms,0,blend_radius_m)
  movel([0.304822, -1.350409, -2.573957, -0.788023, 1.570796, 1.875619],accel_mss,speed_ms,0,blend_radius_m)
  movel([0.304810, -1.350640, -2.573802, -0.787947, 1.570796, 1.875606],accel_mss,speed_ms,0,blend_radius_m)
  movel([0.304780, -1.350876, -2.573644, -0.787869, 1.570796, 1.875576],accel_mss,speed_ms,0,blend_radius_m)
  movel([0.304736, -1.351117, -2.573482, -0.787789, 1.570796, 1.875532],accel_mss,speed_ms,0,blend_radius_m)
  movel([0.304671, -1.351406, -2.573289, -0.787694, 1.570796, 1.875468],accel_mss,speed_ms,0,blend_radius_m)
  movel([0.304594, -1.351698, -2.573093, -0.787598, 1.570796, 1.875391],accel_mss,speed_ms,0,blend_radius_m)
  movel([0.304507, -1.351994, -2.572894, -0.787501, 1.570796, 1.875303],accel_mss,speed_ms,0,blend_radius_m)
  movel([0.304411, -1.352286, -2.572698, -0.787405, 1.570796, 1.875208],accel_mss,speed_ms,0,blend_radius_m)
  movel([0.304305, -1.352581, -2.572500, -0.787308, 1.570796, 1.875102],accel_mss,speed_ms,0,blend_radius_m)
  movel([0.304190, -1.352875, -2.572302, -0.787212, 1.570796, 1.874987],accel_mss,speed_ms,0,blend_radius_m)
  movel([0.304083, -1.353116, -2.572140, -0.787133, 1.570796, 1.874879],accel_mss,speed_ms,0,blend_radius_m)
  movel([0.303962, -1.353358, -2.571977, -0.787054, 1.570796, 1.874758],accel_mss,speed_ms,0,blend_radius_m)
  movel([0.303829, -1.353597, -2.571816, -0.786976, 1.570796, 1.874626],accel_mss,speed_ms,0,blend_radius_m)
  movel([0.303632, -1.353920, -2.571598, -0.786871, 1.570796, 1.874429],accel_mss,speed_ms,0,blend_radius_m)
  movel([0.303419, -1.354237, -2.571384, -0.786768, 1.570796, 1.874215],accel_mss,speed_ms,0,blend_radius_m)
  movel([0.303192, -1.354549, -2.571174, -0.786666, 1.570796, 1.873989],accel_mss,speed_ms,0,blend_radius_m)
  movel([0.302951, -1.354858, -2.570965, -0.786566, 1.570796, 1.873747],accel_mss,speed_ms,0,blend_radius_m)
  movel([0.302696, -1.355159, -2.570761, -0.786468, 1.570796, 1.873492],accel_mss,speed_ms,0,blend_radius_m)
  movel([0.302434, -1.355446, -2.570568, -0.786375, 1.570796, 1.873230],accel_mss,speed_ms,0,blend_radius_m)
  movel([0.302161, -1.355724, -2.570379, -0.786285, 1.570796, 1.872957],accel_mss,speed_ms,0,blend_radius_m)
  movel([0.301874, -1.355993, -2.570197, -0.786198, 1.570796, 1.872671],accel_mss,speed_ms,0,blend_radius_m)
  movel([0.301579, -1.356254, -2.570021, -0.786114, 1.570796, 1.872375],accel_mss,speed_ms,0,blend_radius_m)
  movel([0.301274, -1.356502, -2.569853, -0.786034, 1.570796, 1.872070],accel_mss,speed_ms,0,blend_radius_m)
  movel([0.300964, -1.356735, -2.569695, -0.785959, 1.570796, 1.871761],accel_mss,speed_ms,0,blend_radius_m)
  movel([0.300645, -1.356956, -2.569545, -0.785888, 1.570796, 1.871441],accel_mss,speed_ms,0,blend_radius_m)
  movel([0.300323, -1.357164, -2.569404, -0.785821, 1.570796, 1.871119],accel_mss,speed_ms,0,blend_radius_m)
  movel([0.299992, -1.357357, -2.569273, -0.785759, 1.570796, 1.870788],accel_mss,speed_ms,0,blend_radius_m)
  movel([0.299659, -1.357535, -2.569152, -0.785702, 1.570796, 1.870455],accel_mss,speed_ms,0,blend_radius_m)
  movel([0.299323, -1.357699, -2.569040, -0.785649, 1.570796, 1.870119],accel_mss,speed_ms,0,blend_radius_m)
  movel([0.298983, -1.357849, -2.568939, -0.785601, 1.570796, 1.869779],accel_mss,speed_ms,0,blend_radius_m)
  movel([0.298641, -1.357981, -2.568849, -0.785559, 1.570796, 1.869437],accel_mss,speed_ms,0,blend_radius_m)
  movel([0.298303, -1.358094, -2.568772, -0.785523, 1.570796, 1.869100],accel_mss,speed_ms,0,blend_radius_m)
  movel([0.297963, -1.358195, -2.568703, -0.785491, 1.570796, 1.868759],accel_mss,speed_ms,0,blend_radius_m)
  movel([0.297675, -1.358263, -2.568657, -0.785469, 1.570796, 1.868471],accel_mss,speed_ms,0,blend_radius_m)
  movel([0.297387, -1.358316, -2.568621, -0.785452, 1.570796, 1.868183],accel_mss,speed_ms,0,blend_radius_m)
  movel([0.297107, -1.358352, -2.568597, -0.785440, 1.570796, 1.867903],accel_mss,speed_ms,0,blend_radius_m)
  movel([0.296830, -1.358372, -2.568583, -0.785434, 1.570796, 1.867626],accel_mss,speed_ms,0,blend_radius_m)
  movel([0.296563, -1.358374, -2.568582, -0.785433, 1.570796, 1.867359],accel_mss,speed_ms,0,blend_radius_m)
  movel([0.296302, -1.358359, -2.568592, -0.785438, 1.570796, 1.867098],accel_mss,speed_ms,0,blend_radius_m)
  movel([0.296048, -1.358328, -2.568613, -0.785448, 1.570796, 1.866844],accel_mss,speed_ms,0,blend_radius_m)
  movel([0.295793, -1.358277, -2.568648, -0.785464, 1.570796, 1.866589],accel_mss,speed_ms,0,blend_radius_m)
  movel([0.295549, -1.358214, -2.568691, -0.785485, 1.570796, 1.866346],accel_mss,speed_ms,0,blend_radius_m)
  movel([0.295313, -1.358134, -2.568745, -0.785510, 1.570796, 1.866110],accel_mss,speed_ms,0,blend_radius_m)
  movel([0.295089, -1.358040, -2.568809, -0.785540, 1.570796, 1.865885],accel_mss,speed_ms,0,blend_radius_m)
  movel([0.294878, -1.357931, -2.568883, -0.785575, 1.570796, 1.865675],accel_mss,speed_ms,0,blend_radius_m)
  movel([0.294679, -1.357809, -2.568966, -0.785614, 1.570796, 1.865475],accel_mss,speed_ms,0,blend_radius_m)
  movel([0.294491, -1.357673, -2.569058, -0.785658, 1.570796, 1.865287],accel_mss,speed_ms,0,blend_radius_m)
  movel([0.294312, -1.357515, -2.569165, -0.785708, 1.570796, 1.865108],accel_mss,speed_ms,0,blend_radius_m)
  movel([0.294143, -1.357348, -2.569279, -0.785762, 1.570796, 1.864940],accel_mss,speed_ms,0,blend_radius_m)
  movel([0.293991, -1.357165, -2.569403, -0.785821, 1.570796, 1.864787],accel_mss,speed_ms,0,blend_radius_m)
  movel([0.293854, -1.356972, -2.569534, -0.785883, 1.570796, 1.864650],accel_mss,speed_ms,0,blend_radius_m)
  movel([0.293731, -1.356768, -2.569673, -0.785949, 1.570796, 1.864528],accel_mss,speed_ms,0,blend_radius_m)
  movel([0.293624, -1.356553, -2.569818, -0.786018, 1.570796, 1.864420],accel_mss,speed_ms,0,blend_radius_m)
  movel([0.293532, -1.356327, -2.569971, -0.786090, 1.570796, 1.864328],accel_mss,speed_ms,0,blend_radius_m)
  movel([0.293455, -1.356089, -2.570133, -0.786167, 1.570796, 1.864252],accel_mss,speed_ms,0,blend_radius_m)
  movel([0.293393, -1.355842, -2.570300, -0.786247, 1.570796, 1.864189],accel_mss,speed_ms,0,blend_radius_m)
  movel([0.293350, -1.355586, -2.570473, -0.786330, 1.570796, 1.864146],accel_mss,speed_ms,0,blend_radius_m)
  movel([0.293321, -1.355323, -2.570651, -0.786415, 1.570796, 1.864117],accel_mss,speed_ms,0,blend_radius_m)
  movel([0.293308, -1.355052, -2.570834, -0.786503, 1.570796, 1.864105],accel_mss,speed_ms,0,blend_radius_m)
  movel([0.293312, -1.354775, -2.571021, -0.786593, 1.570796, 1.864108],accel_mss,speed_ms,0,blend_radius_m)
  movel([0.293331, -1.354493, -2.571212, -0.786684, 1.570796, 1.864127],accel_mss,speed_ms,0,blend_radius_m)
  movel([0.293369, -1.354164, -2.571433, -0.786791, 1.570796, 1.864165],accel_mss,speed_ms,0,blend_radius_m)
  movel([0.293421, -1.353831, -2.571658, -0.786900, 1.570796, 1.864217],accel_mss,speed_ms,0,blend_radius_m)
  speed_ms = 0.003
  movel([0.293421, -1.341199, -2.565402, -0.805788, 1.570796, 1.864217],accel_mss,speed_ms,0,blend_radius_m)
  speed_ms = 0.01
  movel([0.293421, -1.317023, -2.552513, -0.842853, 1.570796, 1.864217],accel_mss,speed_ms,0,blend_radius_m)
  movel([0.294198, -1.317224, -2.552384, -0.842780, 1.570796, 1.864995],accel_mss,speed_ms,0,blend_radius_m)
  movel([0.294198, -1.341397, -2.565271, -0.805721, 1.570796, 1.864995],accel_mss,speed_ms,0,blend_radius_m)
  speed_ms = 0.003
  movel([0.294198, -1.350836, -2.569974, -0.791579, 1.570796, 1.864995],accel_mss,speed_ms,0,blend_radius_m)
  speed_ms = 0.007
  movel([0.294328, -1.350403, -2.570264, -0.791722, 1.570796, 1.865125],accel_mss,speed_ms,0,blend_radius_m)
  movel([0.294461, -1.349970, -2.570555, -0.791864, 1.570796, 1.865257],accel_mss,speed_ms,0,blend_radius_m)
  movel([0.294606, -1.349528, -2.570851, -0.792010, 1.570796, 1.865402],accel_mss,speed_ms,0,blend_radius_m)
  movel([0.294752, -1.349088, -2.571145, -0.792156, 1.570796, 1.865549],accel_mss,speed_ms,0,blend_radius_m)
  movel([0.294837, -1.348866, -2.571293, -0.792229, 1.570796, 1.865633],accel_mss,speed_ms,0,blend_radius_m)
  movel([0.294935, -1.348645, -2.571441, -0.792303, 1.570796, 1.865731],accel_mss,speed_ms,0,blend_radius_m)
  movel([0.295004, -1.348518, -2.571526, -0.792345, 1.570796, 1.865800],accel_mss,speed_ms,0,blend_radius_m)
  movel([0.295079, -1.348392, -2.571610, -0.792387, 1.570796, 1.865875],accel_mss,speed_ms,0,blend_radius_m)
  movel([0.295161, -1.348268, -2.571693, -0.792428, 1.570796, 1.865957],accel_mss,speed_ms,0,blend_radius_m)
  movel([0.295358, -1.347996, -2.571874, -0.792518, 1.570796, 1.866154],accel_mss,speed_ms,0,blend_radius_m)
  movel([0.295562, -1.347731, -2.572051, -0.792607, 1.570796, 1.866358],accel_mss,speed_ms,0,blend_radius_m)
  movel([0.295771, -1.347472, -2.572224, -0.792693, 1.570796, 1.866568],accel_mss,speed_ms,0,blend_radius_m)
  movel([0.295993, -1.347218, -2.572393, -0.792778, 1.570796, 1.866790],accel_mss,speed_ms,0,blend_radius_m)
  movel([0.296225, -1.346972, -2.572557, -0.792860, 1.570796, 1.867021],accel_mss,speed_ms,0,blend_radius_m)
  movel([0.296463, -1.346733, -2.572716, -0.792940, 1.570796, 1.867260],accel_mss,speed_ms,0,blend_radius_m)
  movel([0.296712, -1.346501, -2.572871, -0.793017, 1.570796, 1.867508],accel_mss,speed_ms,0,blend_radius_m)
  movel([0.296969, -1.346276, -2.573020, -0.793093, 1.570796, 1.867766],accel_mss,speed_ms,0,blend_radius_m)
  movel([0.297227, -1.346067, -2.573159, -0.793163, 1.570796, 1.868023],accel_mss,speed_ms,0,blend_radius_m)
  movel([0.297491, -1.345867, -2.573292, -0.793230, 1.570796, 1.868288],accel_mss,speed_ms,0,blend_radius_m)
  movel([0.297765, -1.345676, -2.573419, -0.793294, 1.570796, 1.868561],accel_mss,speed_ms,0,blend_radius_m)
  movel([0.298029, -1.345505, -2.573533, -0.793351, 1.570796, 1.868825],accel_mss,speed_ms,0,blend_radius_m)
  movel([0.298297, -1.345344, -2.573639, -0.793405, 1.570796, 1.869094],accel_mss,speed_ms,0,blend_radius_m)
  movel([0.298571, -1.345197, -2.573737, -0.793455, 1.570796, 1.869367],accel_mss,speed_ms,0,blend_radius_m)
  movel([0.298828, -1.345072, -2.573820, -0.793497, 1.570796, 1.869625],accel_mss,speed_ms,0,blend_radius_m)
  movel([0.299083, -1.344954, -2.573898, -0.793537, 1.570796, 1.869879],accel_mss,speed_ms,0,blend_radius_m)
  movel([0.299278, -1.344877, -2.573949, -0.793563, 1.570796, 1.870074],accel_mss,speed_ms,0,blend_radius_m)
  movel([0.299470, -1.344813, -2.573991, -0.793584, 1.570796, 1.870267],accel_mss,speed_ms,0,blend_radius_m)
  movel([0.299688, -1.344761, -2.574026, -0.793602, 1.570796, 1.870484],accel_mss,speed_ms,0,blend_radius_m)
  movel([0.299899, -1.344721, -2.574053, -0.793615, 1.570796, 1.870695],accel_mss,speed_ms,0,blend_radius_m)
  movel([0.300243, -1.344672, -2.574085, -0.793632, 1.570796, 1.871039],accel_mss,speed_ms,0,blend_radius_m)
  movel([0.300586, -1.344630, -2.574113, -0.793646, 1.570796, 1.871383],accel_mss,speed_ms,0,blend_radius_m)
  movel([0.300934, -1.344592, -2.574138, -0.793659, 1.570796, 1.871730],accel_mss,speed_ms,0,blend_radius_m)
  movel([0.301281, -1.344561, -2.574159, -0.793669, 1.570796, 1.872077],accel_mss,speed_ms,0,blend_radius_m)
  movel([0.301481, -1.344554, -2.574163, -0.793672, 1.570796, 1.872278],accel_mss,speed_ms,0,blend_radius_m)
  movel([0.301676, -1.344563, -2.574157, -0.793669, 1.570796, 1.872473],accel_mss,speed_ms,0,blend_radius_m)
  movel([0.301848, -1.344587, -2.574142, -0.793661, 1.570796, 1.872644],accel_mss,speed_ms,0,blend_radius_m)
  movel([0.302010, -1.344627, -2.574115, -0.793647, 1.570796, 1.872806],accel_mss,speed_ms,0,blend_radius_m)
  movel([0.302230, -1.344704, -2.574064, -0.793621, 1.570796, 1.873026],accel_mss,speed_ms,0,blend_radius_m)
  movel([0.302443, -1.344789, -2.574008, -0.793592, 1.570796, 1.873239],accel_mss,speed_ms,0,blend_radius_m)
  movel([0.302651, -1.344890, -2.573941, -0.793558, 1.570796, 1.873447],accel_mss,speed_ms,0,blend_radius_m)
  movel([0.302850, -1.345003, -2.573865, -0.793520, 1.570796, 1.873646],accel_mss,speed_ms,0,blend_radius_m)
  movel([0.303031, -1.345135, -2.573778, -0.793476, 1.570796, 1.873827],accel_mss,speed_ms,0,blend_radius_m)
  movel([0.303198, -1.345279, -2.573682, -0.793427, 1.570796, 1.873995],accel_mss,speed_ms,0,blend_radius_m)
  movel([0.303349, -1.345439, -2.573576, -0.793374, 1.570796, 1.874145],accel_mss,speed_ms,0,blend_radius_m)
  movel([0.303486, -1.345612, -2.573462, -0.793316, 1.570796, 1.874282],accel_mss,speed_ms,0,blend_radius_m)
  movel([0.303608, -1.345802, -2.573335, -0.793252, 1.570796, 1.874404],accel_mss,speed_ms,0,blend_radius_m)
  movel([0.303717, -1.346003, -2.573202, -0.793184, 1.570796, 1.874513],accel_mss,speed_ms,0,blend_radius_m)
  movel([0.303807, -1.346217, -2.573060, -0.793113, 1.570796, 1.874603],accel_mss,speed_ms,0,blend_radius_m)
  movel([0.303883, -1.346439, -2.572912, -0.793038, 1.570796, 1.874679],accel_mss,speed_ms,0,blend_radius_m)
  movel([0.303942, -1.346670, -2.572758, -0.792961, 1.570796, 1.874738],accel_mss,speed_ms,0,blend_radius_m)
  movel([0.303984, -1.346910, -2.572599, -0.792881, 1.570796, 1.874780],accel_mss,speed_ms,0,blend_radius_m)
  movel([0.304009, -1.347163, -2.572430, -0.792796, 1.570796, 1.874806],accel_mss,speed_ms,0,blend_radius_m)
  movel([0.304016, -1.347422, -2.572257, -0.792710, 1.570796, 1.874813],accel_mss,speed_ms,0,blend_radius_m)
  movel([0.304007, -1.347687, -2.572081, -0.792621, 1.570796, 1.874804],accel_mss,speed_ms,0,blend_radius_m)
  movel([0.303980, -1.347959, -2.571899, -0.792531, 1.570796, 1.874776],accel_mss,speed_ms,0,blend_radius_m)
  movel([0.303937, -1.348233, -2.571717, -0.792440, 1.570796, 1.874734],accel_mss,speed_ms,0,blend_radius_m)
  movel([0.303879, -1.348512, -2.571530, -0.792347, 1.570796, 1.874675],accel_mss,speed_ms,0,blend_radius_m)
  movel([0.303801, -1.348794, -2.571342, -0.792254, 1.570796, 1.874598],accel_mss,speed_ms,0,blend_radius_m)
  movel([0.303710, -1.349075, -2.571154, -0.792160, 1.570796, 1.874506],accel_mss,speed_ms,0,blend_radius_m)
  movel([0.303601, -1.349357, -2.570965, -0.792067, 1.570796, 1.874397],accel_mss,speed_ms,0,blend_radius_m)
  movel([0.303476, -1.349641, -2.570775, -0.791973, 1.570796, 1.874272],accel_mss,speed_ms,0,blend_radius_m)
  movel([0.303336, -1.349925, -2.570585, -0.791879, 1.570796, 1.874133],accel_mss,speed_ms,0,blend_radius_m)
  movel([0.303181, -1.350205, -2.570397, -0.791787, 1.570796, 1.873978],accel_mss,speed_ms,0,blend_radius_m)
  movel([0.303018, -1.350476, -2.570216, -0.791698, 1.570796, 1.873815],accel_mss,speed_ms,0,blend_radius_m)
  movel([0.302839, -1.350745, -2.570035, -0.791609, 1.570796, 1.873636],accel_mss,speed_ms,0,blend_radius_m)
  movel([0.302653, -1.351009, -2.569858, -0.791522, 1.570796, 1.873449],accel_mss,speed_ms,0,blend_radius_m)
  movel([0.302453, -1.351269, -2.569683, -0.791437, 1.570796, 1.873250],accel_mss,speed_ms,0,blend_radius_m)
  movel([0.302246, -1.351517, -2.569517, -0.791356, 1.570796, 1.873043],accel_mss,speed_ms,0,blend_radius_m)
  movel([0.302029, -1.351761, -2.569353, -0.791276, 1.570796, 1.872825],accel_mss,speed_ms,0,blend_radius_m)
  movel([0.301802, -1.351997, -2.569194, -0.791198, 1.570796, 1.872599],accel_mss,speed_ms,0,blend_radius_m)
  movel([0.301564, -1.352225, -2.569040, -0.791124, 1.570796, 1.872361],accel_mss,speed_ms,0,blend_radius_m)
  movel([0.301323, -1.352443, -2.568894, -0.791053, 1.570796, 1.872119],accel_mss,speed_ms,0,blend_radius_m)
  movel([0.301073, -1.352652, -2.568753, -0.790984, 1.570796, 1.871869],accel_mss,speed_ms,0,blend_radius_m)
  movel([0.300816, -1.352851, -2.568619, -0.790919, 1.570796, 1.871613],accel_mss,speed_ms,0,blend_radius_m)
  movel([0.300551, -1.353042, -2.568490, -0.790857, 1.570796, 1.871347],accel_mss,speed_ms,0,blend_radius_m)
  movel([0.300280, -1.353223, -2.568368, -0.790798, 1.570796, 1.871076],accel_mss,speed_ms,0,blend_radius_m)
  movel([0.300006, -1.353390, -2.568255, -0.790744, 1.570796, 1.870802],accel_mss,speed_ms,0,blend_radius_m)
  movel([0.299729, -1.353546, -2.568150, -0.790693, 1.570796, 1.870525],accel_mss,speed_ms,0,blend_radius_m)
  movel([0.299446, -1.353692, -2.568051, -0.790646, 1.570796, 1.870242],accel_mss,speed_ms,0,blend_radius_m)
  movel([0.299211, -1.353804, -2.567976, -0.790609, 1.570796, 1.870008],accel_mss,speed_ms,0,blend_radius_m)
  movel([0.298976, -1.353904, -2.567908, -0.790577, 1.570796, 1.869772],accel_mss,speed_ms,0,blend_radius_m)
  movel([0.298781, -1.353977, -2.567859, -0.790553, 1.570796, 1.869578],accel_mss,speed_ms,0,blend_radius_m)
  movel([0.298590, -1.354035, -2.567820, -0.790534, 1.570796, 1.869386],accel_mss,speed_ms,0,blend_radius_m)
  movel([0.298374, -1.354088, -2.567784, -0.790517, 1.570796, 1.869170],accel_mss,speed_ms,0,blend_radius_m)
  movel([0.298159, -1.354126, -2.567758, -0.790505, 1.570796, 1.868955],accel_mss,speed_ms,0,blend_radius_m)
  movel([0.297828, -1.354172, -2.567727, -0.790490, 1.570796, 1.868625],accel_mss,speed_ms,0,blend_radius_m)
  movel([0.297500, -1.354212, -2.567700, -0.790477, 1.570796, 1.868297],accel_mss,speed_ms,0,blend_radius_m)
  movel([0.297176, -1.354246, -2.567677, -0.790466, 1.570796, 1.867972],accel_mss,speed_ms,0,blend_radius_m)
  movel([0.296852, -1.354275, -2.567658, -0.790456, 1.570796, 1.867648],accel_mss,speed_ms,0,blend_radius_m)
  movel([0.296645, -1.354285, -2.567651, -0.790453, 1.570796, 1.867441],accel_mss,speed_ms,0,blend_radius_m)
  movel([0.296449, -1.354278, -2.567655, -0.790455, 1.570796, 1.867245],accel_mss,speed_ms,0,blend_radius_m)
  movel([0.296278, -1.354262, -2.567666, -0.790461, 1.570796, 1.867075],accel_mss,speed_ms,0,blend_radius_m)
  movel([0.296121, -1.354229, -2.567689, -0.790471, 1.570796, 1.866917],accel_mss,speed_ms,0,blend_radius_m)
  movel([0.295935, -1.354174, -2.567726, -0.790489, 1.570796, 1.866731],accel_mss,speed_ms,0,blend_radius_m)
  movel([0.295754, -1.354113, -2.567767, -0.790509, 1.570796, 1.866550],accel_mss,speed_ms,0,blend_radius_m)
  movel([0.295553, -1.354024, -2.567827, -0.790538, 1.570796, 1.866349],accel_mss,speed_ms,0,blend_radius_m)
  movel([0.295368, -1.353920, -2.567897, -0.790571, 1.570796, 1.866165],accel_mss,speed_ms,0,blend_radius_m)
  movel([0.295196, -1.353802, -2.567977, -0.790610, 1.570796, 1.865992],accel_mss,speed_ms,0,blend_radius_m)
  movel([0.295024, -1.353659, -2.568074, -0.790656, 1.570796, 1.865820],accel_mss,speed_ms,0,blend_radius_m)
  movel([0.294865, -1.353503, -2.568179, -0.790707, 1.570796, 1.865661],accel_mss,speed_ms,0,blend_radius_m)
  movel([0.294721, -1.353336, -2.568291, -0.790761, 1.570796, 1.865518],accel_mss,speed_ms,0,blend_radius_m)
  movel([0.294587, -1.353155, -2.568414, -0.790820, 1.570796, 1.865383],accel_mss,speed_ms,0,blend_radius_m)
  movel([0.294469, -1.352961, -2.568544, -0.790883, 1.570796, 1.865265],accel_mss,speed_ms,0,blend_radius_m)
  movel([0.294364, -1.352759, -2.568681, -0.790949, 1.570796, 1.865161],accel_mss,speed_ms,0,blend_radius_m)
  movel([0.294280, -1.352551, -2.568821, -0.791017, 1.570796, 1.865076],accel_mss,speed_ms,0,blend_radius_m)
  movel([0.294210, -1.352336, -2.568966, -0.791087, 1.570796, 1.865007],accel_mss,speed_ms,0,blend_radius_m)
  movel([0.294158, -1.352109, -2.569118, -0.791162, 1.570796, 1.864954],accel_mss,speed_ms,0,blend_radius_m)
  movel([0.294120, -1.351874, -2.569276, -0.791239, 1.570796, 1.864916],accel_mss,speed_ms,0,blend_radius_m)
  movel([0.294091, -1.351633, -2.569438, -0.791317, 1.570796, 1.864887],accel_mss,speed_ms,0,blend_radius_m)
  movel([0.294085, -1.351517, -2.569516, -0.791355, 1.570796, 1.864882],accel_mss,speed_ms,0,blend_radius_m)
  movel([0.294088, -1.351398, -2.569596, -0.791394, 1.570796, 1.864884],accel_mss,speed_ms,0,blend_radius_m)
  movel([0.294101, -1.351276, -2.569679, -0.791435, 1.570796, 1.864897],accel_mss,speed_ms,0,blend_radius_m)
  movel([0.294142, -1.351058, -2.569825, -0.791506, 1.570796, 1.864938],accel_mss,speed_ms,0,blend_radius_m)
  movel([0.294198, -1.350836, -2.569974, -0.791579, 1.570796, 1.864995],accel_mss,speed_ms,0,blend_radius_m)
  speed_ms = 0.003
  movel([0.294198, -1.354028, -2.571525, -0.786836, 1.570796, 1.864995],accel_mss,speed_ms,0,blend_radius_m)
  speed_ms = 0.007
  movel([0.294328, -1.353596, -2.571816, -0.786976, 1.570796, 1.865125],accel_mss,speed_ms,0,blend_radius_m)
  movel([0.294461, -1.353164, -2.572108, -0.787118, 1.570796, 1.865257],accel_mss,speed_ms,0,blend_radius_m)
  movel([0.294606, -1.352723, -2.572404, -0.787262, 1.570796, 1.865402],accel_mss,speed_ms,0,blend_radius_m)
  movel([0.294752, -1.352284, -2.572699, -0.787406, 1.570796, 1.865549],accel_mss,speed_ms,0,blend_radius_m)
  movel([0.294837, -1.352063, -2.572848, -0.787478, 1.570796, 1.865633],accel_mss,speed_ms,0,blend_radius_m)
  movel([0.294935, -1.351843, -2.572996, -0.787551, 1.570796, 1.865731],accel_mss,speed_ms,0,blend_radius_m)
  movel([0.295004, -1.351715, -2.573081, -0.787592, 1.570796, 1.865800],accel_mss,speed_ms,0,blend_radius_m)
  movel([0.295079, -1.351590, -2.573165, -0.787634, 1.570796, 1.865875],accel_mss,speed_ms,0,blend_radius_m)
  movel([0.295161, -1.351465, -2.573249, -0.787675, 1.570796, 1.865957],accel_mss,speed_ms,0,blend_radius_m)
  movel([0.295358, -1.351195, -2.573430, -0.787764, 1.570796, 1.866154],accel_mss,speed_ms,0,blend_radius_m)
  movel([0.295562, -1.350930, -2.573608, -0.787851, 1.570796, 1.866358],accel_mss,speed_ms,0,blend_radius_m)
  movel([0.295771, -1.350672, -2.573781, -0.787936, 1.570796, 1.866568],accel_mss,speed_ms,0,blend_radius_m)
  movel([0.295993, -1.350418, -2.573951, -0.788020, 1.570796, 1.866790],accel_mss,speed_ms,0,blend_radius_m)
  movel([0.296225, -1.350172, -2.574115, -0.788101, 1.570796, 1.867021],accel_mss,speed_ms,0,blend_radius_m)
  movel([0.296463, -1.349935, -2.574274, -0.788180, 1.570796, 1.867260],accel_mss,speed_ms,0,blend_radius_m)
  movel([0.296712, -1.349703, -2.574429, -0.788257, 1.570796, 1.867508],accel_mss,speed_ms,0,blend_radius_m)
  movel([0.296969, -1.349479, -2.574579, -0.788331, 1.570796, 1.867766],accel_mss,speed_ms,0,blend_radius_m)
  movel([0.297227, -1.349270, -2.574718, -0.788401, 1.570796, 1.868023],accel_mss,speed_ms,0,blend_radius_m)
  movel([0.297491, -1.349070, -2.574852, -0.788467, 1.570796, 1.868288],accel_mss,speed_ms,0,blend_radius_m)
  movel([0.297765, -1.348880, -2.574979, -0.788530, 1.570796, 1.868561],accel_mss,speed_ms,0,blend_radius_m)
  movel([0.298029, -1.348709, -2.575093, -0.788587, 1.570796, 1.868825],accel_mss,speed_ms,0,blend_radius_m)
  movel([0.298297, -1.348549, -2.575199, -0.788641, 1.570796, 1.869094],accel_mss,speed_ms,0,blend_radius_m)
  movel([0.298571, -1.348402, -2.575298, -0.788690, 1.570796, 1.869367],accel_mss,speed_ms,0,blend_radius_m)
  movel([0.298828, -1.348277, -2.575381, -0.788731, 1.570796, 1.869625],accel_mss,speed_ms,0,blend_radius_m)
  movel([0.299083, -1.348159, -2.575459, -0.788771, 1.570796, 1.869879],accel_mss,speed_ms,0,blend_radius_m)
  movel([0.299278, -1.348082, -2.575511, -0.788796, 1.570796, 1.870074],accel_mss,speed_ms,0,blend_radius_m)
  movel([0.299470, -1.348019, -2.575553, -0.788817, 1.570796, 1.870267],accel_mss,speed_ms,0,blend_radius_m)
  movel([0.299688, -1.347967, -2.575587, -0.788835, 1.570796, 1.870484],accel_mss,speed_ms,0,blend_radius_m)
  movel([0.299899, -1.347927, -2.575614, -0.788848, 1.570796, 1.870695],accel_mss,speed_ms,0,blend_radius_m)
  movel([0.300243, -1.347878, -2.575647, -0.788864, 1.570796, 1.871039],accel_mss,speed_ms,0,blend_radius_m)
  movel([0.300586, -1.347836, -2.575675, -0.788878, 1.570796, 1.871383],accel_mss,speed_ms,0,blend_radius_m)
  movel([0.300934, -1.347798, -2.575700, -0.788891, 1.570796, 1.871730],accel_mss,speed_ms,0,blend_radius_m)
  movel([0.301281, -1.347767, -2.575720, -0.788901, 1.570796, 1.872077],accel_mss,speed_ms,0,blend_radius_m)
  movel([0.301481, -1.347760, -2.575725, -0.788904, 1.570796, 1.872278],accel_mss,speed_ms,0,blend_radius_m)
  movel([0.301676, -1.347770, -2.575719, -0.788901, 1.570796, 1.872473],accel_mss,speed_ms,0,blend_radius_m)
  movel([0.301848, -1.347793, -2.575703, -0.788893, 1.570796, 1.872644],accel_mss,speed_ms,0,blend_radius_m)
  movel([0.302010, -1.347833, -2.575676, -0.788879, 1.570796, 1.872806],accel_mss,speed_ms,0,blend_radius_m)
  movel([0.302230, -1.347910, -2.575625, -0.788854, 1.570796, 1.873026],accel_mss,speed_ms,0,blend_radius_m)
  movel([0.302443, -1.347995, -2.575569, -0.788825, 1.570796, 1.873239],accel_mss,speed_ms,0,blend_radius_m)
  movel([0.302651, -1.348096, -2.575502, -0.788792, 1.570796, 1.873447],accel_mss,speed_ms,0,blend_radius_m)
  movel([0.302850, -1.348209, -2.575426, -0.788754, 1.570796, 1.873646],accel_mss,speed_ms,0,blend_radius_m)
  movel([0.303031, -1.348340, -2.575339, -0.788710, 1.570796, 1.873827],accel_mss,speed_ms,0,blend_radius_m)
  movel([0.303198, -1.348484, -2.575243, -0.788662, 1.570796, 1.873995],accel_mss,speed_ms,0,blend_radius_m)
  movel([0.303349, -1.348643, -2.575137, -0.788609, 1.570796, 1.874145],accel_mss,speed_ms,0,blend_radius_m)
  movel([0.303486, -1.348816, -2.575022, -0.788552, 1.570796, 1.874282],accel_mss,speed_ms,0,blend_radius_m)
  movel([0.303608, -1.349005, -2.574895, -0.788489, 1.570796, 1.874404],accel_mss,speed_ms,0,blend_radius_m)
  movel([0.303717, -1.349206, -2.574761, -0.788422, 1.570796, 1.874513],accel_mss,speed_ms,0,blend_radius_m)
  movel([0.303807, -1.349419, -2.574619, -0.788351, 1.570796, 1.874603],accel_mss,speed_ms,0,blend_radius_m)
  movel([0.303883, -1.349641, -2.574470, -0.788277, 1.570796, 1.874679],accel_mss,speed_ms,0,blend_radius_m)
  movel([0.303942, -1.349872, -2.574316, -0.788201, 1.570796, 1.874738],accel_mss,speed_ms,0,blend_radius_m)
  movel([0.303984, -1.350111, -2.574156, -0.788122, 1.570796, 1.874780],accel_mss,speed_ms,0,blend_radius_m)
  movel([0.304009, -1.350363, -2.573988, -0.788038, 1.570796, 1.874806],accel_mss,speed_ms,0,blend_radius_m)
